  movel([-0.123614, -0.788371, -2.798725, -1.125292, 1.570796, 1.447182],accel_mss,speed_ms,0,blend_radius_m)
  movel([-0.122358, -0.787472, -2.798871, -1.126045, 1.570796, 1.448438],accel_mss,speed_ms,0,blend_radius_m)
  movel([-0.121105, -0.786979, -2.798951, -1.126459, 1.570796, 1.449692],accel_mss,speed_ms,0,blend_radius_m)
  movel([-0.120159, -0.787158, -2.798922, -1.126309, 1.570796, 1.450637],accel_mss,speed_ms,0,blend_radius_m)
  movel([-0.119008, -0.788690, -2.798674, -1.125025, 1.570796, 1.451789],accel_mss,speed_ms,0,blend_radius_m)
  movel([-0.118135, -0.791492, -2.798216, -1.122680, 1.570796, 1.452661],accel_mss,speed_ms,0,blend_radius_m)
  movel([-0.117601, -0.794594, -2.797706, -1.120090, 1.570796, 1.453195],accel_mss,speed_ms,0,blend_radius_m)
  movel([-0.115239, -0.789926, -2.798473, -1.123991, 1.570796, 1.455558],accel_mss,speed_ms,0,blend_radius_m)
  movel([-0.112520, -0.785198, -2.799238, -1.127953, 1.570796, 1.458276],accel_mss,speed_ms,0,blend_radius_m)
  movel([-0.109499, -0.780473, -2.799992, -1.131924, 1.570796, 1.461298],accel_mss,speed_ms,0,blend_radius_m)
  movel([-0.106241, -0.775820, -2.800723, -1.135846, 1.570796, 1.464556],accel_mss,speed_ms,0,blend_radius_m)
  movel([-0.099689, -0.766469, -2.802160, -1.143759, 1.570796, 1.471108],accel_mss,speed_ms,0,blend_radius_m)
  movel([-0.097728, -0.763893, -2.802549, -1.145948, 1.570796, 1.473068],accel_mss,speed_ms,0,blend_radius_m)
  movel([-0.095794, -0.761589, -2.802893, -1.147907, 1.570796, 1.475003],accel_mss,speed_ms,0,blend_radius_m)
  movel([-0.093954, -0.759736, -2.803169, -1.149484, 1.570796, 1.476842],accel_mss,speed_ms,0,blend_radius_m)
  movel([-0.092299, -0.758522, -2.803348, -1.150519, 1.570796, 1.478498],accel_mss,speed_ms,0,blend_radius_m)
  movel([-0.090884, -0.758158, -2.803402, -1.150829, 1.570796, 1.479912],accel_mss,speed_ms,0,blend_radius_m)
  movel([-0.089878, -0.758679, -2.803325, -1.150385, 1.570796, 1.480919],accel_mss,speed_ms,0,blend_radius_m)
  movel([-0.089251, -0.759892, -2.803145, -1.149351, 1.570796, 1.481545],accel_mss,speed_ms,0,blend_radius_m)
  movel([-0.088991, -0.761609, -2.802890, -1.147890, 1.570796, 1.481805],accel_mss,speed_ms,0,blend_radius_m)
  movel([-0.089073, -0.763633, -2.802588, -1.146168, 1.570796, 1.481724],accel_mss,speed_ms,0,blend_radius_m)
  movel([-0.089471, -0.765770, -2.802266, -1.144353, 1.570796, 1.481326],accel_mss,speed_ms,0,blend_radius_m)
  movel([-0.090165, -0.767829, -2.801954, -1.142606, 1.570796, 1.480631],accel_mss,speed_ms,0,blend_radius_m)
  movel([-0.091138, -0.769624, -2.801680, -1.141085, 1.570796, 1.479658],accel_mss,speed_ms,0,blend_radius_m)
  movel([-0.085055, -0.761341, -2.802930, -1.148118, 1.570796, 1.485742],accel_mss,speed_ms,0,blend_radius_m)
  movel([-0.081792, -0.757306, -2.803527, -1.151555, 1.570796, 1.489004],accel_mss,speed_ms,0,blend_radius_m)
  movel([-0.078396, -0.753391, -2.804099, -1.154899, 1.570796, 1.492400],accel_mss,speed_ms,0,blend_radius_m)
  movel([-0.074888, -0.749633, -2.804641, -1.158115, 1.570796, 1.495909],accel_mss,speed_ms,0,blend_radius_m)
  movel([-0.071275, -0.746070, -2.805148, -1.161171, 1.570796, 1.499521],accel_mss,speed_ms,0,blend_radius_m)
  movel([-0.067576, -0.742740, -2.805617, -1.164032, 1.570796, 1.503221],accel_mss,speed_ms,0,blend_radius_m)
  movel([-0.063806, -0.739679, -2.806043, -1.166667, 1.570796, 1.506991],accel_mss,speed_ms,0,blend_radius_m)
  movel([-0.061242, -0.738118, -2.806259, -1.168012, 1.570796, 1.509554],accel_mss,speed_ms,0,blend_radius_m)
  movel([-0.058496, -0.737145, -2.806393, -1.168852, 1.570796, 1.512301],accel_mss,speed_ms,0,blend_radius_m)
  movel([-0.057304, -0.737032, -2.806408, -1.168948, 1.570796, 1.513493],accel_mss,speed_ms,0,blend_radius_m)
  movel([-0.056360, -0.737246, -2.806379, -1.168764, 1.570796, 1.514437],accel_mss,speed_ms,0,blend_radius_m)
  movel([-0.055759, -0.737845, -2.806297, -1.168247, 1.570796, 1.515037],accel_mss,speed_ms,0,blend_radius_m)
  movel([-0.055607, -0.738896, -2.806152, -1.167342, 1.570796, 1.515190],accel_mss,speed_ms,0,blend_radius_m)
  movel([-0.055970, -0.740265, -2.805962, -1.166162, 1.570796, 1.514827],accel_mss,speed_ms,0,blend_radius_m)
  movel([-0.056714, -0.741799, -2.805748, -1.164841, 1.570796, 1.514083],accel_mss,speed_ms,0,blend_radius_m)
  movel([-0.058927, -0.745239, -2.805266, -1.161885, 1.570796, 1.511869],accel_mss,speed_ms,0,blend_radius_m)
  movel([-0.061573, -0.748454, -2.804809, -1.159126, 1.570796, 1.509223],accel_mss,speed_ms,0,blend_radius_m)
  movel([-0.064470, -0.751417, -2.804384, -1.156588, 1.570796, 1.506326],accel_mss,speed_ms,0,blend_radius_m)
  movel([-0.067437, -0.754102, -2.803995, -1.154291, 1.570796, 1.503359],accel_mss,speed_ms,0,blend_radius_m)
  movel([-0.063607, -0.752594, -2.804214, -1.155581, 1.570796, 1.507189],accel_mss,speed_ms,0,blend_radius_m)
  movel([-0.059620, -0.750631, -2.804497, -1.157260, 1.570796, 1.511176],accel_mss,speed_ms,0,blend_radius_m)
  movel([-0.055519, -0.748238, -2.804840, -1.159311, 1.570796, 1.515278],accel_mss,speed_ms,0,blend_radius_m)
  movel([-0.051338, -0.745435, -2.805238, -1.161716, 1.570796, 1.519459],accel_mss,speed_ms,0,blend_radius_m)
  movel([-0.048030, -0.742875, -2.805598, -1.163916, 1.570796, 1.522766],accel_mss,speed_ms,0,blend_radius_m)
  movel([-0.041537, -0.737330, -2.806367, -1.168691, 1.570796, 1.529259],accel_mss,speed_ms,0,blend_radius_m)
  movel([-0.038202, -0.734723, -2.806724, -1.170942, 1.570796, 1.532595],accel_mss,speed_ms,0,blend_radius_m)
  movel([-0.034400, -0.732028, -2.807090, -1.173271, 1.570796, 1.536396],accel_mss,speed_ms,0,blend_radius_m)
  movel([-0.027997, -0.727831, -2.807652, -1.176906, 1.570796, 1.542799],accel_mss,speed_ms,0,blend_radius_m)
  movel([-0.024935, -0.726094, -2.807883, -1.178413, 1.570796, 1.545861],accel_mss,speed_ms,0,blend_radius_m)
  movel([-0.022568, -0.725095, -2.808015, -1.179280, 1.570796, 1.548229],accel_mss,speed_ms,0,blend_radius_m)
  movel([-0.021784, -0.724985, -2.808029, -1.179375, 1.570796, 1.549013],accel_mss,speed_ms,0,blend_radius_m)
  movel([-0.021347, -0.725203, -2.808001, -1.179186, 1.570796, 1.549449],accel_mss,speed_ms,0,blend_radius_m)
  movel([-0.021306, -0.725781, -2.807924, -1.178683, 1.570796, 1.549490],accel_mss,speed_ms,0,blend_radius_m)
  movel([-0.021722, -0.726772, -2.807793, -1.177824, 1.570796, 1.549074],accel_mss,speed_ms,0,blend_radius_m)
  movel([-0.023301, -0.729254, -2.807462, -1.175672, 1.570796, 1.547495],accel_mss,speed_ms,0,blend_radius_m)
  movel([-0.025347, -0.731856, -2.807113, -1.173420, 1.570796, 1.545450],accel_mss,speed_ms,0,blend_radius_m)
  movel([-0.027725, -0.734514, -2.806753, -1.171123, 1.570796, 1.543072],accel_mss,speed_ms,0,blend_radius_m)
  movel([-0.030292, -0.737144, -2.806393, -1.168852, 1.570796, 1.540504],accel_mss,speed_ms,0,blend_radius_m)
  movel([-0.035478, -0.742049, -2.805713, -1.164626, 1.570796, 1.535318],accel_mss,speed_ms,0,blend_radius_m)
  movel([-0.039835, -0.745995, -2.805159, -1.161235, 1.570796, 1.530962],accel_mss,speed_ms,0,blend_radius_m)
  movel([-0.037640, -0.745598, -2.805215, -1.161576, 1.570796, 1.533156],accel_mss,speed_ms,0,blend_radius_m)
  movel([-0.035326, -0.744930, -2.805309, -1.162150, 1.570796, 1.535470],accel_mss,speed_ms,0,blend_radius_m)
  movel([-0.030418, -0.742923, -2.805591, -1.163875, 1.570796, 1.540378],accel_mss,speed_ms,0,blend_radius_m)
  movel([-0.025249, -0.740229, -2.805967, -1.166193, 1.570796, 1.545548],accel_mss,speed_ms,0,blend_radius_m)
  movel([-0.019955, -0.737110, -2.806398, -1.168881, 1.570796, 1.550841],accel_mss,speed_ms,0,blend_radius_m)
  movel([-0.015550, -0.734257, -2.806788, -1.171345, 1.570796, 1.555246],accel_mss,speed_ms,0,blend_radius_m)
  movel([-0.002182, -0.725105, -2.808013, -1.179270, 1.570796, 1.568614],accel_mss,speed_ms,0,blend_radius_m)
  movel([0.000291, -0.723828, -2.808181, -1.180380, 1.570796, 1.571087],accel_mss,speed_ms,0,blend_radius_m)
  movel([0.002219, -0.723407, -2.808237, -1.180746, 1.570796, 1.573015],accel_mss,speed_ms,0,blend_radius_m)
  movel([0.002614, -0.723722, -2.808195, -1.180471, 1.570796, 1.573410],accel_mss,speed_ms,0,blend_radius_m)
  movel([0.002432, -0.724499, -2.808093, -1.179796, 1.570796, 1.573228],accel_mss,speed_ms,0,blend_radius_m)
  movel([0.001528, -0.725818, -2.807919, -1.178652, 1.570796, 1.572325],accel_mss,speed_ms,0,blend_radius_m)
  movel([-0.000242, -0.727756, -2.807662, -1.176971, 1.570796, 1.570554],accel_mss,speed_ms,0,blend_radius_m)
  movel([-0.003204, -0.730567, -2.807287, -1.174536, 1.570796, 1.567592],accel_mss,speed_ms,0,blend_radius_m)
  movel([-0.006618, -0.733453, -2.806897, -1.172039, 1.570796, 1.564179],accel_mss,speed_ms,0,blend_radius_m)
  movel([-0.009977, -0.735885, -2.806566, -1.169939, 1.570796, 1.560819],accel_mss,speed_ms,0,blend_radius_m)
  movel([-0.011482, -0.736767, -2.806445, -1.169177, 1.570796, 1.559315],accel_mss,speed_ms,0,blend_radius_m)
  movel([-0.012779, -0.737329, -2.806368, -1.168692, 1.570796, 1.558017],accel_mss,speed_ms,0,blend_radius_m)
  movel([-0.007737, -0.737133, -2.806395, -1.168862, 1.570796, 1.563059],accel_mss,speed_ms,0,blend_radius_m)
  movel([-0.002332, -0.736239, -2.806517, -1.169632, 1.570796, 1.568464],accel_mss,speed_ms,0,blend_radius_m)
  movel([0.003362, -0.734781, -2.806716, -1.170892, 1.570796, 1.574158],accel_mss,speed_ms,0,blend_radius_m)
  movel([0.009278, -0.732894, -2.806973, -1.172522, 1.570796, 1.580074],accel_mss,speed_ms,0,blend_radius_m)
  movel([0.021466, -0.728361, -2.807582, -1.176446, 1.570796, 1.592262],accel_mss,speed_ms,0,blend_radius_m)
  movel([0.033600, -0.723736, -2.808193, -1.180459, 1.570796, 1.604396],accel_mss,speed_ms,0,blend_radius_m)
  movel([0.035605, -0.723312, -2.808249, -1.180828, 1.570796, 1.606402],accel_mss,speed_ms,0,blend_radius_m)
  movel([0.036255, -0.723590, -2.808212, -1.180586, 1.570796, 1.607051],accel_mss,speed_ms,0,blend_radius_m)
  movel([0.036422, -0.724403, -2.808106, -1.179880, 1.570796, 1.607218],accel_mss,speed_ms,0,blend_radius_m)
  movel([0.036036, -0.725600, -2.807948, -1.178841, 1.570796, 1.606833],accel_mss,speed_ms,0,blend_radius_m)
  movel([0.034004, -0.728911, -2.807508, -1.175970, 1.570796, 1.604800],accel_mss,speed_ms,0,blend_radius_m)
  movel([0.032557, -0.730811, -2.807254, -1.174324, 1.570796, 1.603354],accel_mss,speed_ms,0,blend_radius_m)
  movel([0.029315, -0.734343, -2.806776, -1.171270, 1.570796, 1.600111],accel_mss,speed_ms,0,blend_radius_m)
  movel([0.025758, -0.737485, -2.806346, -1.168557, 1.570796, 1.596555],accel_mss,speed_ms,0,blend_radius_m)
  movel([0.022037, -0.740240, -2.805965, -1.166184, 1.570796, 1.592834],accel_mss,speed_ms,0,blend_radius_m)
  movel([0.018315, -0.742582, -2.805639, -1.164168, 1.570796, 1.589112],accel_mss,speed_ms,0,blend_radius_m)
  movel([0.014745, -0.744506, -2.805369, -1.162514, 1.570796, 1.585541],accel_mss,speed_ms,0,blend_radius_m)
  movel([0.011481, -0.745991, -2.805159, -1.161239, 1.570796, 1.582277],accel_mss,speed_ms,0,blend_radius_m)
  movel([0.008687, -0.747012, -2.805015, -1.160363, 1.570796, 1.579483],accel_mss,speed_ms,0,blend_radius_m)
  movel([0.008653, -0.747858, -2.804894, -1.159637, 1.570796, 1.579449],accel_mss,speed_ms,0,blend_radius_m)
  movel([0.009139, -0.748262, -2.804836, -1.159290, 1.570796, 1.579935],accel_mss,speed_ms,0,blend_radius_m)
  movel([0.010647, -0.748657, -2.804780, -1.158952, 1.570796, 1.581444],accel_mss,speed_ms,0,blend_radius_m)
  movel([0.012360, -0.748723, -2.804771, -1.158895, 1.570796, 1.583157],accel_mss,speed_ms,0,blend_radius_m)
  movel([0.016128, -0.748272, -2.804835, -1.159282, 1.570796, 1.586925],accel_mss,speed_ms,0,blend_radius_m)
  movel([0.022850, -0.747039, -2.805011, -1.160339, 1.570796, 1.593647],accel_mss,speed_ms,0,blend_radius_m)
  movel([0.029687, -0.745518, -2.805226, -1.161645, 1.570796, 1.600483],accel_mss,speed_ms,0,blend_radius_m)
  movel([0.043712, -0.741725, -2.805759, -1.164905, 1.570796, 1.614508],accel_mss,speed_ms,0,blend_radius_m)
  movel([0.047601, -0.740757, -2.805894, -1.165738, 1.570796, 1.618397],accel_mss,speed_ms,0,blend_radius_m)
  movel([0.050057, -0.740378, -2.805946, -1.166065, 1.570796, 1.620854],accel_mss,speed_ms,0,blend_radius_m)
  movel([0.052405, -0.740305, -2.805956, -1.166128, 1.570796, 1.623201],accel_mss,speed_ms,0,blend_radius_m)
  movel([0.054288, -0.740724, -2.805898, -1.165767, 1.570796, 1.625084],accel_mss,speed_ms,0,blend_radius_m)
  movel([0.055366, -0.741799, -2.805748, -1.164841, 1.570796, 1.626162],accel_mss,speed_ms,0,blend_radius_m)
  movel([0.055503, -0.742631, -2.805632, -1.164126, 1.570796, 1.626300],accel_mss,speed_ms,0,blend_radius_m)
  movel([0.055317, -0.743690, -2.805484, -1.163216, 1.570796, 1.626113],accel_mss,speed_ms,0,blend_radius_m)
  movel([0.054755, -0.745002, -2.805299, -1.162088, 1.570796, 1.625552],accel_mss,speed_ms,0,blend_radius_m)
  movel([0.053791, -0.746577, -2.805076, -1.160736, 1.570796, 1.624588],accel_mss,speed_ms,0,blend_radius_m)
  movel([0.052380, -0.748019, -2.804871, -1.159499, 1.570796, 1.623176],accel_mss,speed_ms,0,blend_radius_m)
  movel([0.050460, -0.749382, -2.804676, -1.158330, 1.570796, 1.621256],accel_mss,speed_ms,0,blend_radius_m)
  movel([0.040183, -0.755535, -2.803787, -1.153068, 1.570796, 1.610979],accel_mss,speed_ms,0,blend_radius_m)
  movel([0.036738, -0.757148, -2.803550, -1.151690, 1.570796, 1.607535],accel_mss,speed_ms,0,blend_radius_m)
  movel([0.035260, -0.757597, -2.803484, -1.151307, 1.570796, 1.606056],accel_mss,speed_ms,0,blend_radius_m)
  movel([0.034042, -0.757700, -2.803469, -1.151220, 1.570796, 1.604838],accel_mss,speed_ms,0,blend_radius_m)
  movel([0.039097, -0.759244, -2.803241, -1.149904, 1.570796, 1.609893],accel_mss,speed_ms,0,blend_radius_m)
  movel([0.044720, -0.759886, -2.803146, -1.149356, 1.570796, 1.615516],accel_mss,speed_ms,0,blend_radius_m)
  movel([0.050778, -0.759793, -2.803160, -1.149436, 1.570796, 1.621574],accel_mss,speed_ms,0,blend_radius_m)
  movel([0.057144, -0.759117, -2.803260, -1.150012, 1.570796, 1.627940],accel_mss,speed_ms,0,blend_radius_m)
  movel([0.062648, -0.757727, -2.803465, -1.151197, 1.570796, 1.633444],accel_mss,speed_ms,0,blend_radius_m)
  movel([0.070534, -0.755900, -2.803733, -1.152756, 1.570796, 1.641330],accel_mss,speed_ms,0,blend_radius_m)
  movel([0.074102, -0.755520, -2.803789, -1.153080, 1.570796, 1.644899],accel_mss,speed_ms,0,blend_radius_m)
  movel([0.076754, -0.755848, -2.803741, -1.152800, 1.570796, 1.647550],accel_mss,speed_ms,0,blend_radius_m)
  movel([0.077577, -0.756361, -2.803666, -1.152363, 1.570796, 1.648374],accel_mss,speed_ms,0,blend_radius_m)
  movel([0.077981, -0.757146, -2.803551, -1.151692, 1.570796, 1.648777],accel_mss,speed_ms,0,blend_radius_m)
  movel([0.077904, -0.758242, -2.803389, -1.150758, 1.570796, 1.648701],accel_mss,speed_ms,0,blend_radius_m)
  movel([0.077296, -0.759666, -2.803179, -1.149544, 1.570796, 1.648093],accel_mss,speed_ms,0,blend_radius_m)
  movel([0.076368, -0.761124, -2.802963, -1.148302, 1.570796, 1.647164],accel_mss,speed_ms,0,blend_radius_m)
  movel([0.075295, -0.762513, -2.802755, -1.147120, 1.570796, 1.646091],accel_mss,speed_ms,0,blend_radius_m)
  movel([0.072924, -0.765097, -2.802368, -1.144925, 1.570796, 1.643720],accel_mss,speed_ms,0,blend_radius_m)
  movel([0.070302, -0.767643, -2.801982, -1.142764, 1.570796, 1.641099],accel_mss,speed_ms,0,blend_radius_m)
  movel([0.064988, -0.772160, -2.801291, -1.138938, 1.570796, 1.635784],accel_mss,speed_ms,0,blend_radius_m)
  movel([0.062326, -0.774111, -2.800989, -1.137289, 1.570796, 1.633122],accel_mss,speed_ms,0,blend_radius_m)
  movel([0.067181, -0.773517, -2.801081, -1.137791, 1.570796, 1.637977],accel_mss,speed_ms,0,blend_radius_m)
  movel([0.072189, -0.772546, -2.801231, -1.138612, 1.570796, 1.642985],accel_mss,speed_ms,0,blend_radius_m)
  movel([0.077338, -0.771243, -2.801432, -1.139714, 1.570796, 1.648134],accel_mss,speed_ms,0,blend_radius_m)
  movel([0.082615, -0.769641, -2.801678, -1.141070, 1.570796, 1.653412],accel_mss,speed_ms,0,blend_radius_m)
  movel([0.093490, -0.765710, -2.802275, -1.144404, 1.570796, 1.664286],accel_mss,speed_ms,0,blend_radius_m)
  movel([0.104701, -0.761055, -2.802973, -1.148361, 1.570796, 1.675497],accel_mss,speed_ms,0,blend_radius_m)
  movel([0.107639, -0.760148, -2.803108, -1.149134, 1.570796, 1.678435],accel_mss,speed_ms,0,blend_radius_m)
  movel([0.108683, -0.760339, -2.803079, -1.148971, 1.570796, 1.679480],accel_mss,speed_ms,0,blend_radius_m)
  movel([0.109107, -0.761285, -2.802939, -1.148165, 1.570796, 1.679903],accel_mss,speed_ms,0,blend_radius_m)
  movel([0.108974, -0.762254, -2.802794, -1.147340, 1.570796, 1.679770],accel_mss,speed_ms,0,blend_radius_m)
  movel([0.108569, -0.763342, -2.802631, -1.146416, 1.570796, 1.679365],accel_mss,speed_ms,0,blend_radius_m)
  movel([0.107060, -0.765815, -2.802259, -1.144315, 1.570796, 1.677856],accel_mss,speed_ms,0,blend_radius_m)
  movel([0.104857, -0.768511, -2.801850, -1.142028, 1.570796, 1.675653],accel_mss,speed_ms,0,blend_radius_m)
  movel([0.102226, -0.771265, -2.801429, -1.139696, 1.570796, 1.673022],accel_mss,speed_ms,0,blend_radius_m)
  movel([0.096762, -0.776227, -2.800659, -1.135502, 1.570796, 1.667558],accel_mss,speed_ms,0,blend_radius_m)
  movel([0.092780, -0.779303, -2.800177, -1.132910, 1.570796, 1.663577],accel_mss,speed_ms,0,blend_radius_m)
  movel([0.095018, -0.778629, -2.800283, -1.133477, 1.570796, 1.665815],accel_mss,speed_ms,0,blend_radius_m)
  movel([0.097342, -0.777697, -2.800429, -1.134262, 1.570796, 1.668138],accel_mss,speed_ms,0,blend_radius_m)
  movel([0.102193, -0.775141, -2.800829, -1.136419, 1.570796, 1.672990],accel_mss,speed_ms,0,blend_radius_m)
  movel([0.107238, -0.771741, -2.801355, -1.139293, 1.570796, 1.678035],accel_mss,speed_ms,0,blend_radius_m)
  movel([0.112383, -0.767625, -2.801985, -1.142779, 1.570796, 1.683179],accel_mss,speed_ms,0,blend_radius_m)
  movel([0.117534, -0.762890, -2.802699, -1.146800, 1.570796, 1.688330],accel_mss,speed_ms,0,blend_radius_m)
  movel([0.122590, -0.757669, -2.803474, -1.151246, 1.570796, 1.693387],accel_mss,speed_ms,0,blend_radius_m)
  movel([0.127452, -0.752066, -2.804291, -1.156033, 1.570796, 1.698249],accel_mss,speed_ms,0,blend_radius_m)
  movel([0.132018, -0.746209, -2.805128, -1.161051, 1.570796, 1.702814],accel_mss,speed_ms,0,blend_radius_m)
  movel([0.134037, -0.743591, -2.805498, -1.163300, 1.570796, 1.704834],accel_mss,speed_ms,0,blend_radius_m)
  movel([0.135120, -0.742450, -2.805657, -1.164281, 1.570796, 1.705916],accel_mss,speed_ms,0,blend_radius_m)
  movel([0.136237, -0.741570, -2.805780, -1.165038, 1.570796, 1.707033],accel_mss,speed_ms,0,blend_radius_m)
  movel([0.137379, -0.741088, -2.805848, -1.165453, 1.570796, 1.708175],accel_mss,speed_ms,0,blend_radius_m)
  movel([0.138333, -0.741050, -2.805853, -1.165486, 1.570796, 1.709129],accel_mss,speed_ms,0,blend_radius_m)
  movel([0.139345, -0.741714, -2.805760, -1.164914, 1.570796, 1.710141],accel_mss,speed_ms,0,blend_radius_m)
  movel([0.139829, -0.743141, -2.805561, -1.163688, 1.570796, 1.710625],accel_mss,speed_ms,0,blend_radius_m)
  movel([0.139879, -0.745135, -2.805280, -1.161974, 1.570796, 1.710675],accel_mss,speed_ms,0,blend_radius_m)
  movel([0.139591, -0.747520, -2.804942, -1.159927, 1.570796, 1.710387],accel_mss,speed_ms,0,blend_radius_m)
  movel([0.138373, -0.752698, -2.804199, -1.155492, 1.570796, 1.709169],accel_mss,speed_ms,0,blend_radius_m)
  movel([0.136926, -0.757207, -2.803542, -1.151641, 1.570796, 1.707723],accel_mss,speed_ms,0,blend_radius_m)
  movel([0.140852, -0.751503, -2.804372, -1.156514, 1.570796, 1.711648],accel_mss,speed_ms,0,blend_radius_m)
  movel([0.144402, -0.745687, -2.805202, -1.161500, 1.570796, 1.715198],accel_mss,speed_ms,0,blend_radius_m)
  movel([0.147549, -0.739819, -2.806024, -1.166546, 1.570796, 1.718345],accel_mss,speed_ms,0,blend_radius_m)
  movel([0.150273, -0.733978, -2.806826, -1.171585, 1.570796, 1.721070],accel_mss,speed_ms,0,blend_radius_m)
  movel([0.152533, -0.728242, -2.807598, -1.176549, 1.570796, 1.723330],accel_mss,speed_ms,0,blend_radius_m)
  movel([0.154318, -0.722674, -2.808332, -1.181382, 1.570796, 1.725114],accel_mss,speed_ms,0,blend_radius_m)
  movel([0.155580, -0.717372, -2.809019, -1.185998, 1.570796, 1.726376],accel_mss,speed_ms,0,blend_radius_m)
  movel([0.156297, -0.712407, -2.809651, -1.190332, 1.570796, 1.727094],accel_mss,speed_ms,0,blend_radius_m)
  movel([0.156402, -0.706121, -2.810434, -1.195834, 1.570796, 1.727198],accel_mss,speed_ms,0,blend_radius_m)
  movel([0.156716, -0.702641, -2.810860, -1.198888, 1.570796, 1.727512],accel_mss,speed_ms,0,blend_radius_m)
  movel([0.157110, -0.700860, -2.811076, -1.200453, 1.570796, 1.727906],accel_mss,speed_ms,0,blend_radius_m)
  movel([0.157721, -0.699072, -2.811292, -1.202026, 1.570796, 1.728517],accel_mss,speed_ms,0,blend_radius_m)
  movel([0.159157, -0.696129, -2.811643, -1.204617, 1.570796, 1.729953],accel_mss,speed_ms,0,blend_radius_m)
  movel([0.160486, -0.694322, -2.811857, -1.206209, 1.570796, 1.731283],accel_mss,speed_ms,0,blend_radius_m)
  movel([0.161725, -0.693413, -2.811965, -1.207012, 1.570796, 1.732521],accel_mss,speed_ms,0,blend_radius_m)
  movel([0.162880, -0.693157, -2.811995, -1.207237, 1.570796, 1.733676],accel_mss,speed_ms,0,blend_radius_m)
  movel([0.165920, -0.693920, -2.811905, -1.206564, 1.570796, 1.736716],accel_mss,speed_ms,0,blend_radius_m)
  movel([0.166833, -0.693867, -2.811911, -1.206611, 1.570796, 1.737629],accel_mss,speed_ms,0,blend_radius_m)
  movel([0.168876, -0.689499, -2.812422, -1.210468, 1.570796, 1.739672],accel_mss,speed_ms,0,blend_radius_m)
  movel([0.170617, -0.685171, -2.812919, -1.214299, 1.570796, 1.741413],accel_mss,speed_ms,0,blend_radius_m)
  movel([0.172069, -0.680901, -2.813402, -1.218086, 1.570796, 1.742866],accel_mss,speed_ms,0,blend_radius_m)
  movel([0.173248, -0.676699, -2.813870, -1.221820, 1.570796, 1.744044],accel_mss,speed_ms,0,blend_radius_m)
  movel([0.174153, -0.672593, -2.814320, -1.225476, 1.570796, 1.744950],accel_mss,speed_ms,0,blend_radius_m)
  movel([0.174801, -0.668595, -2.814751, -1.229043, 1.570796, 1.745598],accel_mss,speed_ms,0,blend_radius_m)
  movel([0.175391, -0.660973, -2.815554, -1.235862, 1.570796, 1.746188],accel_mss,speed_ms,0,blend_radius_m)
  movel([0.175103, -0.653985, -2.816269, -1.242134, 1.570796, 1.745899],accel_mss,speed_ms,0,blend_radius_m)
  movel([0.174059, -0.647747, -2.816891, -1.247751, 1.570796, 1.744855],accel_mss,speed_ms,0,blend_radius_m)
  movel([0.172351, -0.642405, -2.817410, -1.252574, 1.570796, 1.743147],accel_mss,speed_ms,0,blend_radius_m)
  movel([0.170116, -0.638064, -2.817824, -1.256502, 1.570796, 1.740912],accel_mss,speed_ms,0,blend_radius_m)
  speed_ms = 0.005
  movel([0.170116, -0.631907, -2.811057, -1.269425, 1.570796, 1.740912],accel_mss,speed_ms,0,blend_radius_m)
  speed_ms = 0.040
  movel([0.138700, -0.656581, -2.808612, -1.247195, 1.570796, 1.709497],accel_mss,speed_ms,0,blend_radius_m)
  speed_ms = 0.005
  movel([0.138700, -0.663123, -2.815330, -1.233936, 1.570796, 1.709497],accel_mss,speed_ms,0,blend_radius_m)
  speed_ms = 0.025
  movel([0.136102, -0.662756, -2.815369, -1.234264, 1.570796, 1.706899],accel_mss,speed_ms,0,blend_radius_m)
  movel([0.133054, -0.663285, -2.815313, -1.233791, 1.570796, 1.703850],accel_mss,speed_ms,0,blend_radius_m)
  movel([0.129644, -0.664578, -2.815178, -1.232634, 1.570796, 1.700441],accel_mss,speed_ms,0,blend_radius_m)
  movel([0.125976, -0.666489, -2.814975, -1.230924, 1.570796, 1.696772],accel_mss,speed_ms,0,blend_radius_m)
  movel([0.122143, -0.668882, -2.814720, -1.228787, 1.570796, 1.692939],accel_mss,speed_ms,0,blend_radius_m)
  movel([0.118234, -0.671617, -2.814426, -1.226346, 1.570796, 1.689030],accel_mss,speed_ms,0,blend_radius_m)
  movel([0.110564, -0.677562, -2.813775, -1.221052, 1.570796, 1.681360],accel_mss,speed_ms,0,blend_radius_m)
  speed_ms = 0.005
  movel([0.110564, -0.670808, -2.807087, -1.234494, 1.570796, 1.681360],accel_mss,speed_ms,0,blend_radius_m)
  speed_ms = 0.040
  movel([0.120496, -0.662365, -2.808003, -1.242021, 1.570796, 1.691293],accel_mss,speed_ms,0,blend_radius_m)
  speed_ms = 0.005
  movel([0.120496, -0.668994, -2.814708, -1.228687, 1.570796, 1.691293],accel_mss,speed_ms,0,blend_radius_m)
  speed_ms = 0.025
  movel([0.122110, -0.664213, -2.815216, -1.232960, 1.570796, 1.692907],accel_mss,speed_ms,0,blend_radius_m)
  movel([0.123299, -0.659769, -2.815679, -1.236941, 1.570796, 1.694095],accel_mss,speed_ms,0,blend_radius_m)
  movel([0.124068, -0.655656, -2.816100, -1.240632, 1.570796, 1.694864],accel_mss,speed_ms,0,blend_radius_m)
  movel([0.124435, -0.651859, -2.816483, -1.244047, 1.570796, 1.695231],accel_mss,speed_ms,0,blend_radius_m)
  movel([0.124423, -0.648357, -2.816831, -1.247202, 1.570796, 1.695219],accel_mss,speed_ms,0,blend_radius_m)
  movel([0.124046, -0.645138, -2.817146, -1.250105, 1.570796, 1.694842],accel_mss,speed_ms,0,blend_radius_m)
  movel([0.123323, -0.642185, -2.817431, -1.252773, 1.570796, 1.694119],accel_mss,speed_ms,0,blend_radius_m)
  movel([0.122274, -0.639481, -2.817690, -1.255219, 1.570796, 1.693071],accel_mss,speed_ms,0,blend_radius_m)
  movel([0.118229, -0.632565, -2.818336, -1.261487, 1.570796, 1.689025],accel_mss,speed_ms,0,blend_radius_m)
  movel([0.116481, -0.629055, -2.818657, -1.264676, 1.570796, 1.687277],accel_mss,speed_ms,0,blend_radius_m)
  movel([0.115290, -0.624496, -2.819067, -1.268826, 1.570796, 1.686086],accel_mss,speed_ms,0,blend_radius_m)
  movel([0.114590, -0.618038, -2.819633, -1.274718, 1.570796, 1.685386],accel_mss,speed_ms,0,blend_radius_m)
  movel([0.114549, -0.610974, -2.820233, -1.281182, 1.570796, 1.685345],accel_mss,speed_ms,0,blend_radius_m)
  movel([0.115398, -0.603180, -2.820873, -1.288336, 1.570796, 1.686195],accel_mss,speed_ms,0,blend_radius_m)
  movel([0.116229, -0.598970, -2.821209, -1.292210, 1.570796, 1.687025],accel_mss,speed_ms,0,blend_radius_m)
  movel([0.117376, -0.594532, -2.821555, -1.296302, 1.570796, 1.688172],accel_mss,speed_ms,0,blend_radius_m)
  movel([0.119840, -0.587296, -2.822104, -1.302989, 1.570796, 1.690636],accel_mss,speed_ms,0,blend_radius_m)
  movel([0.123098, -0.579856, -2.822647, -1.309886, 1.570796, 1.693894],accel_mss,speed_ms,0,blend_radius_m)
  movel([0.127112, -0.572263, -2.823180, -1.316946, 1.570796, 1.697908],accel_mss,speed_ms,0,blend_radius_m)
  movel([0.131842, -0.564581, -2.823697, -1.324111, 1.570796, 1.702638],accel_mss,speed_ms,0,blend_radius_m)
  movel([0.137234, -0.556886, -2.824193, -1.331309, 1.570796, 1.708030],accel_mss,speed_ms,0,blend_radius_m)
  movel([0.143247, -0.549247, -2.824664, -1.338478, 1.570796, 1.714044],accel_mss,speed_ms,0,blend_radius_m)
  movel([0.149829, -0.541732, -2.825106, -1.345550, 1.570796, 1.720625],accel_mss,speed_ms,0,blend_radius_m)
  movel([0.156913, -0.534435, -2.825516, -1.352438, 1.570796, 1.727709],accel_mss,speed_ms,0,blend_radius_m)
  movel([0.162439, -0.529240, -2.825796, -1.357352, 1.570796, 1.733235],accel_mss,speed_ms,0,blend_radius_m)
  movel([0.168059, -0.524374, -2.826050, -1.361965, 1.570796, 1.738855],accel_mss,speed_ms,0,blend_radius_m)
  movel([0.173713, -0.519879, -2.826276, -1.366234, 1.570796, 1.744510],accel_mss,speed_ms,0,blend_radius_m)
  movel([0.179359, -0.515772, -2.826477, -1.370140, 1.570796, 1.750155],accel_mss,speed_ms,0,blend_radius_m)
  movel([0.184932, -0.512108, -2.826651, -1.373629, 1.570796, 1.755728],accel_mss,speed_ms,0,blend_radius_m)
  movel([0.190379, -0.508915, -2.826799, -1.376675, 1.570796, 1.761175],accel_mss,speed_ms,0,blend_radius_m)
  movel([0.195640, -0.506227, -2.826921, -1.379241, 1.570796, 1.766437],accel_mss,speed_ms,0,blend_radius_m)
  movel([0.200660, -0.504082, -2.827016, -1.381291, 1.570796, 1.771456],accel_mss,speed_ms,0,blend_radius_m)
  movel([0.205378, -0.502513, -2.827085, -1.382791, 1.570796, 1.776175],accel_mss,speed_ms,0,blend_radius_m)
  movel([0.209750, -0.501543, -2.827127, -1.383719, 1.570796, 1.780546],accel_mss,speed_ms,0,blend_radius_m)
  movel([0.213716, -0.501208, -2.827141, -1.384040, 1.570796, 1.784512],accel_mss,speed_ms,0,blend_radius_m)
  movel([0.217226, -0.501531, -2.827127, -1.383731, 1.570796, 1.788023],accel_mss,speed_ms,0,blend_radius_m)
  movel([0.220235, -0.502533, -2.827084, -1.382772, 1.570796, 1.791031],accel_mss,speed_ms,0,blend_radius_m)
  movel([0.222682, -0.504249, -2.827009, -1.381132, 1.570796, 1.793478],accel_mss,speed_ms,0,blend_radius_m)
  movel([0.224532, -0.506682, -2.826900, -1.378807, 1.570796, 1.795329],accel_mss,speed_ms,0,blend_radius_m)
  movel([0.225745, -0.509859, -2.826756, -1.375774, 1.570796, 1.796541],accel_mss,speed_ms,0,blend_radius_m)
  movel([0.226531, -0.514797, -2.826524, -1.371068, 1.570796, 1.797328],accel_mss,speed_ms,0,blend_radius_m)
  movel([0.226728, -0.520288, -2.826256, -1.365845, 1.570796, 1.797524],accel_mss,speed_ms,0,blend_radius_m)
  movel([0.226455, -0.526200, -2.825956, -1.360233, 1.570796, 1.797251],accel_mss,speed_ms,0,blend_radius_m)
  movel([0.225856, -0.532375, -2.825628, -1.354386, 1.570796, 1.796653],accel_mss,speed_ms,0,blend_radius_m)
  movel([0.223911, -0.546253, -2.824843, -1.341294, 1.570796, 1.794707],accel_mss,speed_ms,0,blend_radius_m)
  movel([0.221348, -0.560558, -2.823959, -1.327872, 1.570796, 1.792145],accel_mss,speed_ms,0,blend_radius_m)
  movel([0.218336, -0.575144, -2.822980, -1.314265, 1.570796, 1.789132],accel_mss,speed_ms,0,blend_radius_m)
  movel([0.215033, -0.589850, -2.821912, -1.300626, 1.570796, 1.785830],accel_mss,speed_ms,0,blend_radius_m)
  movel([0.201838, -0.647356, -2.816929, -1.248104, 1.570796, 1.772635],accel_mss,speed_ms,0,blend_radius_m)
  movel([0.196552, -0.674366, -2.814127, -1.223896, 1.570796, 1.767348],accel_mss,speed_ms,0,blend_radius_m)
  movel([0.194383, -0.687392, -2.812665, -1.212332, 1.570796, 1.765179],accel_mss,speed_ms,0,blend_radius_m)
  movel([0.192649, -0.699989, -2.811181, -1.201218, 1.570796, 1.763445],accel_mss,speed_ms,0,blend_radius_m)
  movel([0.191422, -0.712103, -2.809689, -1.190597, 1.570796, 1.762219],accel_mss,speed_ms,0,blend_radius_m)
  movel([0.190783, -0.723666, -2.808203, -1.180520, 1.570796, 1.761579],accel_mss,speed_ms,0,blend_radius_m)
  movel([0.190794, -0.734632, -2.806737, -1.171020, 1.570796, 1.761590],accel_mss,speed_ms,0,blend_radius_m)
  movel([0.191537, -0.744943, -2.805307, -1.162139, 1.570796, 1.762333],accel_mss,speed_ms,0,blend_radius_m)
  movel([0.192118, -0.748698, -2.804774, -1.158917, 1.570796, 1.762914],accel_mss,speed_ms,0,blend_radius_m)
  movel([0.193186, -0.751978, -2.804303, -1.156107, 1.570796, 1.763982],accel_mss,speed_ms,0,blend_radius_m)
  movel([0.194999, -0.754344, -2.803960, -1.154085, 1.570796, 1.765795],accel_mss,speed_ms,0,blend_radius_m)
  movel([0.196267, -0.755045, -2.803858, -1.153486, 1.570796, 1.767064],accel_mss,speed_ms,0,blend_radius_m)
  movel([0.197826, -0.755346, -2.803814, -1.153229, 1.570796, 1.768623],accel_mss,speed_ms,0,blend_radius_m)
  speed_ms = 0.005
  movel([0.197826, -0.747557, -2.797313, -1.167520, 1.570796, 1.768623],accel_mss,speed_ms,0,blend_radius_m)
  speed_ms = 0.040
  movel([0.166317, -0.709653, -2.802474, -1.200262, 1.570796, 1.737113],accel_mss,speed_ms,0,blend_radius_m)
  speed_ms = 0.005
  movel([0.166317, -0.716956, -2.809072, -1.186361, 1.570796, 1.737113],accel_mss,speed_ms,0,blend_radius_m)
  speed_ms = 0.025
  movel([0.165098, -0.718894, -2.808823, -1.184672, 1.570796, 1.735894],accel_mss,speed_ms,0,blend_radius_m)
  movel([0.164169, -0.720873, -2.808567, -1.182949, 1.570796, 1.734965],accel_mss,speed_ms,0,blend_radius_m)
  movel([0.163511, -0.722861, -2.808308, -1.181220, 1.570796, 1.734307],accel_mss,speed_ms,0,blend_radius_m)
  movel([0.163074, -0.724875, -2.808044, -1.179471, 1.570796, 1.733870],accel_mss,speed_ms,0,blend_radius_m)
  movel([0.162764, -0.728898, -2.807510, -1.175981, 1.570796, 1.733560],accel_mss,speed_ms,0,blend_radius_m)
  movel([0.162975, -0.732871, -2.806976, -1.172543, 1.570796, 1.733771],accel_mss,speed_ms,0,blend_radius_m)
  movel([0.164204, -0.743735, -2.805477, -1.163177, 1.570796, 1.735001],accel_mss,speed_ms,0,blend_radius_m)
  movel([0.163980, -0.746745, -2.805052, -1.160591, 1.570796, 1.734776],accel_mss,speed_ms,0,blend_radius_m)
  movel([0.163462, -0.748245, -2.804839, -1.159305, 1.570796, 1.734258],accel_mss,speed_ms,0,blend_radius_m)
  movel([0.162572, -0.749528, -2.804656, -1.158205, 1.570796, 1.733369],accel_mss,speed_ms,0,blend_radius_m)
  movel([0.161731, -0.750298, -2.804545, -1.157545, 1.570796, 1.732527],accel_mss,speed_ms,0,blend_radius_m)
  movel([0.160936, -0.750613, -2.804500, -1.157276, 1.570796, 1.731733],accel_mss,speed_ms,0,blend_radius_m)
  movel([0.160186, -0.750538, -2.804511, -1.157340, 1.570796, 1.730982],accel_mss,speed_ms,0,blend_radius_m)
  movel([0.158834, -0.749419, -2.804671, -1.158299, 1.570796, 1.729630],accel_mss,speed_ms,0,blend_radius_m)
  movel([0.157687, -0.747402, -2.804959, -1.160028, 1.570796, 1.728483],accel_mss,speed_ms,0,blend_radius_m)
  movel([0.156071, -0.742470, -2.805655, -1.164264, 1.570796, 1.726867],accel_mss,speed_ms,0,blend_radius_m)
  movel([0.155517, -0.739344, -2.806090, -1.166956, 1.570796, 1.726314],accel_mss,speed_ms,0,blend_radius_m)
  movel([0.153840, -0.744960, -2.805305, -1.162125, 1.570796, 1.724636],accel_mss,speed_ms,0,blend_radius_m)
  movel([0.152864, -0.750190, -2.804561, -1.157639, 1.570796, 1.723661],accel_mss,speed_ms,0,blend_radius_m)
  movel([0.152485, -0.755065, -2.803855, -1.153468, 1.570796, 1.723281],accel_mss,speed_ms,0,blend_radius_m)
  movel([0.152612, -0.759591, -2.803190, -1.149608, 1.570796, 1.723409],accel_mss,speed_ms,0,blend_radius_m)
  movel([0.153139, -0.763802, -2.802562, -1.146024, 1.570796, 1.723935],accel_mss,speed_ms,0,blend_radius_m)
  movel([0.153986, -0.767697, -2.801974, -1.142718, 1.570796, 1.724782],accel_mss,speed_ms,0,blend_radius_m)
  movel([0.156246, -0.774616, -2.800910, -1.136862, 1.570796, 1.727042],accel_mss,speed_ms,0,blend_radius_m)
  movel([0.156304, -0.776266, -2.800653, -1.135470, 1.570796, 1.727100],accel_mss,speed_ms,0,blend_radius_m)
  movel([0.155931, -0.777204, -2.800507, -1.134678, 1.570796, 1.726728],accel_mss,speed_ms,0,blend_radius_m)
  movel([0.155223, -0.778000, -2.800382, -1.134007, 1.570796, 1.726019],accel_mss,speed_ms,0,blend_radius_m)
  movel([0.154317, -0.778384, -2.800321, -1.133684, 1.570796, 1.725113],accel_mss,speed_ms,0,blend_radius_m)
  movel([0.152367, -0.778552, -2.800295, -1.133542, 1.570796, 1.723163],accel_mss,speed_ms,0,blend_radius_m)
  movel([0.150735, -0.778213, -2.800348, -1.133827, 1.570796, 1.721532],accel_mss,speed_ms,0,blend_radius_m)
  movel([0.149384, -0.777445, -2.800469, -1.134475, 1.570796, 1.720180],accel_mss,speed_ms,0,blend_radius_m)
  movel([0.148290, -0.776299, -2.800648, -1.135442, 1.570796, 1.719086],accel_mss,speed_ms,0,blend_radius_m)
  movel([0.146758, -0.773161, -2.801136, -1.138092, 1.570796, 1.717554],accel_mss,speed_ms,0,blend_radius_m)
  movel([0.145914, -0.769328, -2.801725, -1.141336, 1.570796, 1.716710],accel_mss,speed_ms,0,blend_radius_m)
  movel([0.145148, -0.778136, -2.800360, -1.133893, 1.570796, 1.715944],accel_mss,speed_ms,0,blend_radius_m)
  movel([0.145196, -0.782168, -2.799723, -1.130499, 1.570796, 1.715993],accel_mss,speed_ms,0,blend_radius_m)
  movel([0.145776, -0.785782, -2.799144, -1.127463, 1.570796, 1.716573],accel_mss,speed_ms,0,blend_radius_m)
  movel([0.146955, -0.788308, -2.798736, -1.125345, 1.570796, 1.717752],accel_mss,speed_ms,0,blend_radius_m)
  movel([0.150125, -0.792178, -2.798104, -1.122107, 1.570796, 1.720921],accel_mss,speed_ms,0,blend_radius_m)
  movel([0.151210, -0.794682, -2.797691, -1.120016, 1.570796, 1.722006],accel_mss,speed_ms,0,blend_radius_m)
  movel([0.151294, -0.795308, -2.797587, -1.119493, 1.570796, 1.722090],accel_mss,speed_ms,0,blend_radius_m)
  movel([0.151105, -0.796095, -2.797457, -1.118837, 1.570796, 1.721902],accel_mss,speed_ms,0,blend_radius_m)
  movel([0.150490, -0.796935, -2.797317, -1.118137, 1.570796, 1.721287],accel_mss,speed_ms,0,blend_radius_m)
  movel([0.149467, -0.797739, -2.797183, -1.117467, 1.570796, 1.720263],accel_mss,speed_ms,0,blend_radius_m)
  movel([0.146733, -0.799179, -2.796941, -1.116269, 1.570796, 1.717529],accel_mss,speed_ms,0,blend_radius_m)
  movel([0.142223, -0.800846, -2.796661, -1.114882, 1.570796, 1.713020],accel_mss,speed_ms,0,blend_radius_m)
  movel([0.142758, -0.803053, -2.796287, -1.113049, 1.570796, 1.713554],accel_mss,speed_ms,0,blend_radius_m)
  movel([0.143619, -0.805415, -2.795885, -1.111089, 1.570796, 1.714415],accel_mss,speed_ms,0,blend_radius_m)
  movel([0.144902, -0.807761, -2.795482, -1.109146, 1.570796, 1.715698],accel_mss,speed_ms,0,blend_radius_m)
  movel([0.146705, -0.809923, -2.795108, -1.107358, 1.570796, 1.717501],accel_mss,speed_ms,0,blend_radius_m)
  movel([0.152042, -0.812028, -2.794742, -1.105619, 1.570796, 1.722838],accel_mss,speed_ms,0,blend_radius_m)
  movel([0.154980, -0.813362, -2.794508, -1.104519, 1.570796, 1.725776],accel_mss,speed_ms,0,blend_radius_m)
  movel([0.155811, -0.814073, -2.794384, -1.103932, 1.570796, 1.726607],accel_mss,speed_ms,0,blend_radius_m)
  movel([0.155954, -0.814801, -2.794255, -1.103332, 1.570796, 1.726751],accel_mss,speed_ms,0,blend_radius_m)
  movel([0.155514, -0.815661, -2.794104, -1.102624, 1.570796, 1.726310],accel_mss,speed_ms,0,blend_radius_m)
  movel([0.154880, -0.816481, -2.793959, -1.101949, 1.570796, 1.725676],accel_mss,speed_ms,0,blend_radius_m)
  movel([0.153372, -0.817748, -2.793735, -1.100907, 1.570796, 1.724168],accel_mss,speed_ms,0,blend_radius_m)
  movel([0.152148, -0.818307, -2.793635, -1.100447, 1.570796, 1.722944],accel_mss,speed_ms,0,blend_radius_m)
  movel([0.150940, -0.818620, -2.793579, -1.100190, 1.570796, 1.721736],accel_mss,speed_ms,0,blend_radius_m)
  movel([0.148664, -0.819018, -2.793508, -1.099862, 1.570796, 1.719461],accel_mss,speed_ms,0,blend_radius_m)
  movel([0.149487, -0.821978, -2.792978, -1.097433, 1.570796, 1.720283],accel_mss,speed_ms,0,blend_radius_m)
  movel([0.150580, -0.824668, -2.792492, -1.095228, 1.570796, 1.721377],accel_mss,speed_ms,0,blend_radius_m)
  movel([0.151941, -0.827078, -2.792054, -1.093257, 1.570796, 1.722738],accel_mss,speed_ms,0,blend_radius_m)
  movel([0.153547, -0.829212, -2.791663, -1.091514, 1.570796, 1.724344],accel_mss,speed_ms,0,blend_radius_m)
  movel([0.155518, -0.830855, -2.791360, -1.090174, 1.570796, 1.726315],accel_mss,speed_ms,0,blend_radius_m)
  movel([0.157892, -0.831960, -2.791156, -1.089273, 1.570796, 1.728688],accel_mss,speed_ms,0,blend_radius_m)
  movel([0.163164, -0.833388, -2.790891, -1.088110, 1.570796, 1.733961],accel_mss,speed_ms,0,blend_radius_m)
  movel([0.164477, -0.834123, -2.790754, -1.087512, 1.570796, 1.735273],accel_mss,speed_ms,0,blend_radius_m)
  movel([0.164731, -0.834865, -2.790615, -1.086908, 1.570796, 1.735527],accel_mss,speed_ms,0,blend_radius_m)
  movel([0.164486, -0.835941, -2.790414, -1.086034, 1.570796, 1.735282],accel_mss,speed_ms,0,blend_radius_m)
  movel([0.163859, -0.836981, -2.790219, -1.085189, 1.570796, 1.734656],accel_mss,speed_ms,0,blend_radius_m)
  movel([0.163012, -0.837903, -2.790045, -1.084441, 1.570796, 1.733808],accel_mss,speed_ms,0,blend_radius_m)
  movel([0.161071, -0.839356, -2.789770, -1.083263, 1.570796, 1.731867],accel_mss,speed_ms,0,blend_radius_m)
  movel([0.158538, -0.840756, -2.789505, -1.082128, 1.570796, 1.729334],accel_mss,speed_ms,0,blend_radius_m)
  movel([0.156117, -0.841803, -2.789305, -1.081281, 1.570796, 1.726913],accel_mss,speed_ms,0,blend_radius_m)
  movel([0.153793, -0.842552, -2.789162, -1.080675, 1.570796, 1.724589],accel_mss,speed_ms,0,blend_radius_m)
  movel([0.151559, -0.843038, -2.789069, -1.080282, 1.570796, 1.722355],accel_mss,speed_ms,0,blend_radius_m)
  movel([0.152827, -0.845070, -2.788679, -1.078639, 1.570796, 1.723624],accel_mss,speed_ms,0,blend_radius_m)
  movel([0.154404, -0.846724, -2.788360, -1.077305, 1.570796, 1.725200],accel_mss,speed_ms,0,blend_radius_m)
  movel([0.156283, -0.847956, -2.788121, -1.076312, 1.570796, 1.727080],accel_mss,speed_ms,0,blend_radius_m)
  movel([0.158458, -0.848729, -2.787971, -1.075689, 1.570796, 1.729255],accel_mss,speed_ms,0,blend_radius_m)
  movel([0.160934, -0.848998, -2.787919, -1.075472, 1.570796, 1.731730],accel_mss,speed_ms,0,blend_radius_m)
  movel([0.163710, -0.848723, -2.787972, -1.075694, 1.570796, 1.734507],accel_mss,speed_ms,0,blend_radius_m)
  movel([0.166787, -0.847855, -2.788141, -1.076393, 1.570796, 1.737583],accel_mss,speed_ms,0,blend_radius_m)
  movel([0.170171, -0.846352, -2.788432, -1.077605, 1.570796, 1.740967],accel_mss,speed_ms,0,blend_radius_m)
  speed_ms = 0.005
  movel([0.170171, -0.837613, -2.782198, -1.092579, 1.570796, 1.740967],accel_mss,speed_ms,0,blend_radius_m)
  speed_ms = 0.040
  movel([0.185325, -0.814540, -2.786475, -1.111374, 1.570796, 1.756121],accel_mss,speed_ms,0,blend_radius_m)
  speed_ms = 0.005
  movel([0.185325, -0.823064, -2.792783, -1.096542, 1.570796, 1.756121],accel_mss,speed_ms,0,blend_radius_m)
  speed_ms = 0.025
  movel([0.179130, -0.822911, -2.792810, -1.096668, 1.570796, 1.749926],accel_mss,speed_ms,0,blend_radius_m)
  movel([0.176504, -0.822539, -2.792877, -1.096973, 1.570796, 1.747300],accel_mss,speed_ms,0,blend_radius_m)
  movel([0.174175, -0.821867, -2.792998, -1.097524, 1.570796, 1.744971],accel_mss,speed_ms,0,blend_radius_m)
  movel([0.172123, -0.820815, -2.793187, -1.098387, 1.570796, 1.742919],accel_mss,speed_ms,0,blend_radius_m)
  movel([0.170335, -0.819304, -2.793457, -1.099628, 1.570796, 1.741131],accel_mss,speed_ms,0,blend_radius_m)
  movel([0.168788, -0.817262, -2.793821, -1.101306, 1.570796, 1.739584],accel_mss,speed_ms,0,blend_radius_m)
  movel([0.167475, -0.814605, -2.794290, -1.103494, 1.570796, 1.738271],accel_mss,speed_ms,0,blend_radius_m)
  movel([0.165467, -0.808324, -2.795385, -1.108681, 1.570796, 1.736263],accel_mss,speed_ms,0,blend_radius_m)
  movel([0.164156, -0.801360, -2.796574, -1.114455, 1.570796, 1.734952],accel_mss,speed_ms,0,blend_radius_m)
  movel([0.163481, -0.793797, -2.797837, -1.120755, 1.570796, 1.734277],accel_mss,speed_ms,0,blend_radius_m)
  movel([0.163370, -0.785739, -2.799151, -1.127499, 1.570796, 1.734166],accel_mss,speed_ms,0,blend_radius_m)
  movel([0.163693, -0.778798, -2.800256, -1.133335, 1.570796, 1.734489],accel_mss,speed_ms,0,blend_radius_m)
  movel([0.164351, -0.771584, -2.801380, -1.139426, 1.570796, 1.735147],accel_mss,speed_ms,0,blend_radius_m)
  movel([0.166427, -0.756480, -2.803648, -1.152261, 1.570796, 1.737223],accel_mss,speed_ms,0,blend_radius_m)
  movel([0.175526, -0.702006, -2.810937, -1.199445, 1.570796, 1.746322],accel_mss,speed_ms,0,blend_radius_m)
  movel([0.177448, -0.690287, -2.812330, -1.209772, 1.570796, 1.748244],accel_mss,speed_ms,0,blend_radius_m)
  movel([0.179180, -0.678587, -2.813661, -1.220141, 1.570796, 1.749976],accel_mss,speed_ms,0,blend_radius_m)
  movel([0.180554, -0.667081, -2.814913, -1.230395, 1.570796, 1.751350],accel_mss,speed_ms,0,blend_radius_m)
  movel([0.181390, -0.655935, -2.816072, -1.240382, 1.570796, 1.752186],accel_mss,speed_ms,0,blend_radius_m)
  movel([0.181508, -0.645334, -2.817127, -1.249928, 1.570796, 1.752305],accel_mss,speed_ms,0,blend_radius_m)
  movel([0.180716, -0.635477, -2.818066, -1.258846, 1.570796, 1.751512],accel_mss,speed_ms,0,blend_radius_m)
  movel([0.179492, -0.628855, -2.818676, -1.264858, 1.570796, 1.750288],accel_mss,speed_ms,0,blend_radius_m)
  movel([0.177674, -0.622575, -2.819237, -1.270577, 1.570796, 1.748470],accel_mss,speed_ms,0,blend_radius_m)
  movel([0.175212, -0.616814, -2.819738, -1.275836, 1.570796, 1.746008],accel_mss,speed_ms,0,blend_radius_m)
  movel([0.172054, -0.611754, -2.820168, -1.280467, 1.570796, 1.742851],accel_mss,speed_ms,0,blend_radius_m)
  movel([0.168163, -0.607565, -2.820516, -1.284308, 1.570796, 1.738959],accel_mss,speed_ms,0,blend_radius_m)
  movel([0.163499, -0.604415, -2.820773, -1.287201, 1.570796, 1.734295],accel_mss,speed_ms,0,blend_radius_m)
  movel([0.158021, -0.602490, -2.820928, -1.288971, 1.570796, 1.728817],accel_mss,speed_ms,0,blend_radius_m)
  movel([0.151716, -0.601943, -2.820972, -1.289473, 1.570796, 1.722513],accel_mss,speed_ms,0,blend_radius_m)
  movel([0.148431, -0.602267, -2.820946, -1.289176, 1.570796, 1.719227],accel_mss,speed_ms,0,blend_radius_m)
  movel([0.144882, -0.603048, -2.820884, -1.288457, 1.570796, 1.715678],accel_mss,speed_ms,0,blend_radius_m)
  movel([0.141095, -0.604309, -2.820782, -1.287298, 1.570796, 1.711892],accel_mss,speed_ms,0,blend_radius_m)
  movel([0.137112, -0.606061, -2.820639, -1.285689, 1.570796, 1.707908],accel_mss,speed_ms,0,blend_radius_m)
  movel([0.132975, -0.608300, -2.820455, -1.283634, 1.570796, 1.703772],accel_mss,speed_ms,0,blend_radius_m)
  movel([0.128708, -0.611053, -2.820227, -1.281110, 1.570796, 1.699505],accel_mss,speed_ms,0,blend_radius_m)
  movel([0.124362, -0.614309, -2.819952, -1.278128, 1.570796, 1.695159],accel_mss,speed_ms,0,blend_radius_m)
  movel([0.119974, -0.618083, -2.819629, -1.274677, 1.570796, 1.690770],accel_mss,speed_ms,0,blend_radius_m)
  speed_ms = 0.005
  movel([0.119974, -0.612246, -2.812827, -1.287316, 1.570796, 1.690770],accel_mss,speed_ms,0,blend_radius_m)
  speed_ms = 0.040
  movel([0.105668, -0.599555, -2.813887, -1.298947, 1.570796, 1.676464],accel_mss,speed_ms,0,blend_radius_m)
  speed_ms = 0.005
  movel([0.105668, -0.605180, -2.820711, -1.286498, 1.570796, 1.676464],accel_mss,speed_ms,0,blend_radius_m)
  speed_ms = 0.025
  movel([0.105208, -0.602800, -2.820903, -1.288686, 1.570796, 1.676004],accel_mss,speed_ms,0,blend_radius_m)
  movel([0.105101, -0.600110, -2.821118, -1.291161, 1.570796, 1.675897],accel_mss,speed_ms,0,blend_radius_m)
  movel([0.105749, -0.594005, -2.821596, -1.296788, 1.570796, 1.676545],accel_mss,speed_ms,0,blend_radius_m)
  movel([0.107230, -0.587216, -2.822110, -1.303063, 1.570796, 1.678026],accel_mss,speed_ms,0,blend_radius_m)
  movel([0.109136, -0.580136, -2.822627, -1.309626, 1.570796, 1.679932],accel_mss,speed_ms,0,blend_radius_m)
  speed_ms = 0.005
  movel([0.109136, -0.574935, -2.815764, -1.321690, 1.570796, 1.679932],accel_mss,speed_ms,0,blend_radius_m)
  speed_ms = 0.040
  movel([0.118580, -0.571553, -2.816004, -1.324833, 1.570796, 1.689376],accel_mss,speed_ms,0,blend_radius_m)
  speed_ms = 0.005
  movel([0.118580, -0.576694, -2.822872, -1.312823, 1.570796, 1.689376],accel_mss,speed_ms,0,blend_radius_m)
  speed_ms = 0.025
  movel([0.117402, -0.575267, -2.822972, -1.314150, 1.570796, 1.688198],accel_mss,speed_ms,0,blend_radius_m)
  movel([0.116582, -0.573518, -2.823093, -1.315777, 1.570796, 1.687379],accel_mss,speed_ms,0,blend_radius_m)
  movel([0.115918, -0.569140, -2.823393, -1.319856, 1.570796, 1.686715],accel_mss,speed_ms,0,blend_radius_m)
  movel([0.116427, -0.563751, -2.823752, -1.324886, 1.570796, 1.687223],accel_mss,speed_ms,0,blend_radius_m)
  movel([0.117944, -0.557530, -2.824152, -1.330706, 1.570796, 1.688741],accel_mss,speed_ms,0,blend_radius_m)
  movel([0.120304, -0.550672, -2.824578, -1.337139, 1.570796, 1.691100],accel_mss,speed_ms,0,blend_radius_m)
  movel([0.123332, -0.543377, -2.825011, -1.344000, 1.570796, 1.694129],accel_mss,speed_ms,0,blend_radius_m)
  movel([0.126853, -0.535849, -2.825438, -1.351102, 1.570796, 1.697649],accel_mss,speed_ms,0,blend_radius_m)
  movel([0.130680, -0.528304, -2.825846, -1.358240, 1.570796, 1.701476],accel_mss,speed_ms,0,blend_radius_m)
  speed_ms = 0.005
  movel([0.130680, -0.524028, -2.818917, -1.369444, 1.570796, 1.701476],accel_mss,speed_ms,0,blend_radius_m)
  speed_ms = 0.040
  movel([0.181260, -0.453275, -2.821737, -1.437377, 1.570796, 1.752057],accel_mss,speed_ms,0,blend_radius_m)
  speed_ms = 0.005
  movel([0.181260, -0.456170, -2.828726, -1.427493, 1.570796, 1.752057],accel_mss,speed_ms,0,blend_radius_m)
  speed_ms = 0.025
  movel([0.176078, -0.462124, -2.828557, -1.421708, 1.570796, 1.746874],accel_mss,speed_ms,0,blend_radius_m)
  movel([0.170926, -0.468393, -2.828365, -1.415631, 1.570796, 1.741722],accel_mss,speed_ms,0,blend_radius_m)
  movel([0.165890, -0.474874, -2.828153, -1.409362, 1.570796, 1.736686],accel_mss,speed_ms,0,blend_radius_m)
  movel([0.161028, -0.481494, -2.827921, -1.402974, 1.570796, 1.731824],accel_mss,speed_ms,0,blend_radius_m)
  movel([0.156423, -0.488161, -2.827672, -1.396555, 1.570796, 1.727219],accel_mss,speed_ms,0,blend_radius_m)
  movel([0.152136, -0.494789, -2.827410, -1.390190, 1.570796, 1.722932],accel_mss,speed_ms,0,blend_radius_m)
  movel([0.148234, -0.501305, -2.827137, -1.383947, 1.570796, 1.719030],accel_mss,speed_ms,0,blend_radius_m)
  movel([0.144778, -0.507634, -2.826857, -1.377898, 1.570796, 1.715575],accel_mss,speed_ms,0,blend_radius_m)
  movel([0.141828, -0.513689, -2.826577, -1.372124, 1.570796, 1.712624],accel_mss,speed_ms,0,blend_radius_m)
  movel([0.139435, -0.519412, -2.826300, -1.366678, 1.570796, 1.710232],accel_mss,speed_ms,0,blend_radius_m)
  movel([0.137657, -0.524728, -2.826032, -1.361629, 1.570796, 1.708453],accel_mss,speed_ms,0,blend_radius_m)
  movel([0.136544, -0.529571, -2.825779, -1.357039, 1.570796, 1.707340],accel_mss,speed_ms,0,blend_radius_m)
  movel([0.136155, -0.533872, -2.825547, -1.352970, 1.570796, 1.706952],accel_mss,speed_ms,0,blend_radius_m)
  movel([0.136543, -0.537565, -2.825343, -1.349481, 1.570796, 1.707339],accel_mss,speed_ms,0,blend_radius_m)
  movel([0.137752, -0.540595, -2.825171, -1.346623, 1.570796, 1.708548],accel_mss,speed_ms,0,blend_radius_m)
  movel([0.139843, -0.542894, -2.825039, -1.344456, 1.570796, 1.710639],accel_mss,speed_ms,0,blend_radius_m)
  speed_ms = 0.005
  movel([0.139843, -0.538352, -2.818127, -1.355910, 1.570796, 1.710639],accel_mss,speed_ms,0,blend_radius_m)
  speed_ms = 0.040
  movel([0.162855, -0.512881, -2.819479, -1.380028, 1.570796, 1.733652],accel_mss,speed_ms,0,blend_radius_m)
  speed_ms = 0.005
  movel([0.162855, -0.516946, -2.826420, -1.369023, 1.570796, 1.733652],accel_mss,speed_ms,0,blend_radius_m)
  speed_ms = 0.025
  movel([0.162384, -0.514031, -2.826561, -1.371797, 1.570796, 1.733180],accel_mss,speed_ms,0,blend_radius_m)
  movel([0.162288, -0.510755, -2.826714, -1.374920, 1.570796, 1.733084],accel_mss,speed_ms,0,blend_radius_m)
  movel([0.162565, -0.507153, -2.826879, -1.378357, 1.570796, 1.733362],accel_mss,speed_ms,0,blend_radius_m)
  movel([0.163216, -0.503245, -2.827053, -1.382092, 1.570796, 1.734012],accel_mss,speed_ms,0,blend_radius_m)
  movel([0.164233, -0.499067, -2.827232, -1.386090, 1.570796, 1.735029],accel_mss,speed_ms,0,blend_radius_m)
  movel([0.165623, -0.494639, -2.827416, -1.390334, 1.570796, 1.736419],accel_mss,speed_ms,0,blend_radius_m)
  movel([0.167387, -0.489981, -2.827602, -1.394806, 1.570796, 1.738183],accel_mss,speed_ms,0,blend_radius_m)
  movel([0.169516, -0.485137, -2.827787, -1.399465, 1.570796, 1.740313],accel_mss,speed_ms,0,blend_radius_m)
  movel([0.172012, -0.480127, -2.827970, -1.404292, 1.570796, 1.742809],accel_mss,speed_ms,0,blend_radius_m)
  movel([0.174881, -0.474973, -2.828149, -1.409266, 1.570796, 1.745678],accel_mss,speed_ms,0,blend_radius_m)
  movel([0.178106, -0.469729, -2.828322, -1.414338, 1.570796, 1.748902],accel_mss,speed_ms,0,blend_radius_m)
  movel([0.181701, -0.464399, -2.828489, -1.419501, 1.570796, 1.752497],accel_mss,speed_ms,0,blend_radius_m)
  movel([0.185655, -0.459027, -2.828646, -1.424716, 1.570796, 1.756451],accel_mss,speed_ms,0,blend_radius_m)
  movel([0.189965, -0.453644, -2.828794, -1.429951, 1.570796, 1.760761],accel_mss,speed_ms,0,blend_radius_m)
  movel([0.194624, -0.448291, -2.828932, -1.435166, 1.570796, 1.765421],accel_mss,speed_ms,0,blend_radius_m)
  movel([0.199621, -0.443002, -2.829058, -1.440329, 1.570796, 1.770417],accel_mss,speed_ms,0,blend_radius_m)
  movel([0.204634, -0.438137, -2.829166, -1.445086, 1.570796, 1.775430],accel_mss,speed_ms,0,blend_radius_m)
  movel([0.209620, -0.433721, -2.829257, -1.449411, 1.570796, 1.780416],accel_mss,speed_ms,0,blend_radius_m)
  movel([0.214539, -0.429759, -2.829333, -1.453297, 1.570796, 1.785336],accel_mss,speed_ms,0,blend_radius_m)
  movel([0.219373, -0.426252, -2.829395, -1.456741, 1.570796, 1.790170],accel_mss,speed_ms,0,blend_radius_m)
  movel([0.224084, -0.423203, -2.829447, -1.459739, 1.570796, 1.794880],accel_mss,speed_ms,0,blend_radius_m)
  movel([0.228628, -0.420629, -2.829488, -1.462273, 1.570796, 1.799425],accel_mss,speed_ms,0,blend_radius_m)
  movel([0.232995, -0.418506, -2.829520, -1.464364, 1.570796, 1.803792],accel_mss,speed_ms,0,blend_radius_m)
  movel([0.237129, -0.416859, -2.829543, -1.465986, 1.570796, 1.807925],accel_mss,speed_ms,0,blend_radius_m)
  movel([0.241016, -0.415678, -2.829560, -1.467151, 1.570796, 1.811812],accel_mss,speed_ms,0,blend_radius_m)
  movel([0.247935, -0.414689, -2.829573, -1.468127, 1.570796, 1.818732],accel_mss,speed_ms,0,blend_radius_m)
  movel([0.250900, -0.414885, -2.829571, -1.467933, 1.570796, 1.821697],accel_mss,speed_ms,0,blend_radius_m)
  movel([0.255753, -0.416602, -2.829547, -1.466240, 1.570796, 1.826549],accel_mss,speed_ms,0,blend_radius_m)
  movel([0.257590, -0.418106, -2.829525, -1.464758, 1.570796, 1.828387],accel_mss,speed_ms,0,blend_radius_m)
  movel([0.259001, -0.420034, -2.829497, -1.462858, 1.570796, 1.829798],accel_mss,speed_ms,0,blend_radius_m)
  speed_ms = 0.005
  movel([0.259001, -0.417864, -2.822491, -1.472034, 1.570796, 1.829798],accel_mss,speed_ms,0,blend_radius_m)
  speed_ms = 0.040
  movel([0.274724, -0.430831, -2.822265, -1.459293, 1.570796, 1.845520],accel_mss,speed_ms,0,blend_radius_m)
  speed_ms = 0.005
  movel([0.274724, -0.433269, -2.829266, -1.449855, 1.570796, 1.845520],accel_mss,speed_ms,0,blend_radius_m)
  speed_ms = 0.025
  movel([0.272812, -0.430079, -2.829327, -1.452983, 1.570796, 1.843609],accel_mss,speed_ms,0,blend_radius_m)
  movel([0.269936, -0.428053, -2.829364, -1.454972, 1.570796, 1.840732],accel_mss,speed_ms,0,blend_radius_m)
  movel([0.266170, -0.427187, -2.829379, -1.455823, 1.570796, 1.836967],accel_mss,speed_ms,0,blend_radius_m)
  movel([0.261578, -0.427480, -2.829374, -1.455536, 1.570796, 1.832374],accel_mss,speed_ms,0,blend_radius_m)
  movel([0.256264, -0.428903, -2.829348, -1.454138, 1.570796, 1.827060],accel_mss,speed_ms,0,blend_radius_m)
  movel([0.250302, -0.431450, -2.829301, -1.451639, 1.570796, 1.821099],accel_mss,speed_ms,0,blend_radius_m)
  movel([0.243802, -0.435085, -2.829229, -1.448075, 1.570796, 1.814599],accel_mss,speed_ms,0,blend_radius_m)
  movel([0.236850, -0.439782, -2.829130, -1.443477, 1.570796, 1.807647],accel_mss,speed_ms,0,blend_radius_m)
  movel([0.229570, -0.445491, -2.829000, -1.437898, 1.570796, 1.800366],accel_mss,speed_ms,0,blend_radius_m)
  movel([0.222137, -0.452098, -2.828835, -1.431456, 1.570796, 1.792933],accel_mss,speed_ms,0,blend_radius_m)
  movel([0.214847, -0.459360, -2.828637, -1.424392, 1.570796, 1.785644],accel_mss,speed_ms,0,blend_radius_m)
  movel([0.208004, -0.467046, -2.828407, -1.416936, 1.570796, 1.778801],accel_mss,speed_ms,0,blend_radius_m)
  movel([0.201871, -0.474943, -2.828150, -1.409295, 1.570796, 1.772667],accel_mss,speed_ms,0,blend_radius_m)
  movel([0.199162, -0.478898, -2.828014, -1.405477, 1.570796, 1.769958],accel_mss,speed_ms,0,blend_radius_m)
  movel([0.196726, -0.482824, -2.827873, -1.401692, 1.570796, 1.767523],accel_mss,speed_ms,0,blend_radius_m)
  movel([0.194595, -0.486701, -2.827728, -1.397960, 1.570796, 1.765391],accel_mss,speed_ms,0,blend_radius_m)
  movel([0.192805, -0.490505, -2.827581, -1.394302, 1.570796, 1.763601],accel_mss,speed_ms,0,blend_radius_m)
  movel([0.191376, -0.494210, -2.827433, -1.390745, 1.570796, 1.762173],accel_mss,speed_ms,0,blend_radius_m)
  movel([0.190353, -0.497782, -2.827286, -1.387320, 1.570796, 1.761149],accel_mss,speed_ms,0,blend_radius_m)
  speed_ms = 0.005
  movel([0.190353, -0.494079, -2.820327, -1.397982, 1.570796, 1.761149],accel_mss,speed_ms,0,blend_radius_m)
  speed_ms = 0.040
  movel([0.225557, -0.482976, -2.820769, -1.408644, 1.570796, 1.796354],accel_mss,speed_ms,0,blend_radius_m)
  speed_ms = 0.005
  movel([0.225557, -0.486462, -2.827737, -1.398189, 1.570796, 1.796354],accel_mss,speed_ms,0,blend_radius_m)
  speed_ms = 0.025
  movel([0.230532, -0.480919, -2.827942, -1.403528, 1.570796, 1.801329],accel_mss,speed_ms,0,blend_radius_m)
  movel([0.235675, -0.475846, -2.828120, -1.408423, 1.570796, 1.806472],accel_mss,speed_ms,0,blend_radius_m)
  movel([0.240904, -0.471270, -2.828273, -1.412847, 1.570796, 1.811700],accel_mss,speed_ms,0,blend_radius_m)
  movel([0.246113, -0.467241, -2.828401, -1.416747, 1.570796, 1.816909],accel_mss,speed_ms,0,blend_radius_m)
  movel([0.251210, -0.463791, -2.828507, -1.420091, 1.570796, 1.822007],accel_mss,speed_ms,0,blend_radius_m)
  movel([0.256093, -0.460955, -2.828591, -1.422843, 1.570796, 1.826889],accel_mss,speed_ms,0,blend_radius_m)
  movel([0.260676, -0.458762, -2.828654, -1.424974, 1.570796, 1.831472],accel_mss,speed_ms,0,blend_radius_m)
  movel([0.264851, -0.457246, -2.828696, -1.426447, 1.570796, 1.835647],accel_mss,speed_ms,0,blend_radius_m)
  movel([0.269216, -0.456489, -2.828717, -1.427183, 1.570796, 1.840012],accel_mss,speed_ms,0,blend_radius_m)
  movel([0.272323, -0.457089, -2.828701, -1.426599, 1.570796, 1.843120],accel_mss,speed_ms,0,blend_radius_m)
  movel([0.274310, -0.458896, -2.828650, -1.424843, 1.570796, 1.845106],accel_mss,speed_ms,0,blend_radius_m)
  movel([0.275291, -0.461777, -2.828567, -1.422045, 1.570796, 1.846087],accel_mss,speed_ms,0,blend_radius_m)
  movel([0.275404, -0.465568, -2.828453, -1.418368, 1.570796, 1.846201],accel_mss,speed_ms,0,blend_radius_m)
  movel([0.274782, -0.470132, -2.828309, -1.413947, 1.570796, 1.845579],accel_mss,speed_ms,0,blend_radius_m)
  movel([0.273555, -0.475317, -2.828138, -1.408934, 1.570796, 1.844351],accel_mss,speed_ms,0,blend_radius_m)
  movel([0.271863, -0.480972, -2.827940, -1.403477, 1.570796, 1.842660],accel_mss,speed_ms,0,blend_radius_m)
  speed_ms = 0.005
  movel([0.271863, -0.477592, -2.820967, -1.413830, 1.570796, 1.842660],accel_mss,speed_ms,0,blend_radius_m)
  speed_ms = 0.040
  movel([0.237934, -0.497934, -2.820164, -1.394291, 1.570796, 1.808730],accel_mss,speed_ms,0,blend_radius_m)
  speed_ms = 0.005
  movel([0.237934, -0.501712, -2.827119, -1.383558, 1.570796, 1.808730],accel_mss,speed_ms,0,blend_radius_m)
  speed_ms = 0.025
  movel([0.242451, -0.499306, -2.827222, -1.385861, 1.570796, 1.813247],accel_mss,speed_ms,0,blend_radius_m)
  movel([0.246530, -0.497618, -2.827293, -1.387478, 1.570796, 1.817326],accel_mss,speed_ms,0,blend_radius_m)
  movel([0.250167, -0.496633, -2.827334, -1.388422, 1.570796, 1.820964],accel_mss,speed_ms,0,blend_radius_m)
  movel([0.253371, -0.496299, -2.827348, -1.388742, 1.570796, 1.824168],accel_mss,speed_ms,0,blend_radius_m)
  movel([0.256145, -0.496592, -2.827336, -1.388461, 1.570796, 1.826941],accel_mss,speed_ms,0,blend_radius_m)
  movel([0.258492, -0.497468, -2.827299, -1.387621, 1.570796, 1.829288],accel_mss,speed_ms,0,blend_radius_m)
  movel([0.260428, -0.498888, -2.827240, -1.386261, 1.570796, 1.831224],accel_mss,speed_ms,0,blend_radius_m)
  movel([0.261949, -0.500825, -2.827158, -1.384407, 1.570796, 1.832745],accel_mss,speed_ms,0,blend_radius_m)
  movel([0.263082, -0.503224, -2.827054, -1.382112, 1.570796, 1.833878],accel_mss,speed_ms,0,blend_radius_m)
  movel([0.263834, -0.506045, -2.826929, -1.379415, 1.570796, 1.834630],accel_mss,speed_ms,0,blend_radius_m)
  movel([0.264212, -0.509256, -2.826784, -1.376350, 1.570796, 1.835008],accel_mss,speed_ms,0,blend_radius_m)
  movel([0.264237, -0.512805, -2.826619, -1.372966, 1.570796, 1.835033],accel_mss,speed_ms,0,blend_radius_m)
  movel([0.263917, -0.516659, -2.826434, -1.369296, 1.570796, 1.834713],accel_mss,speed_ms,0,blend_radius_m)
  movel([0.262305, -0.525101, -2.826012, -1.361276, 1.570796, 1.833101],accel_mss,speed_ms,0,blend_radius_m)
  movel([0.261033, -0.529618, -2.825776, -1.356995, 1.570796, 1.831830],accel_mss,speed_ms,0,blend_radius_m)
  movel([0.260911, -0.528484, -2.825836, -1.358069, 1.570796, 1.831708],accel_mss,speed_ms,0,blend_radius_m)
  speed_ms = 0.005
  movel([0.260911, -0.524205, -2.818907, -1.369276, 1.570796, 1.831708],accel_mss,speed_ms,0,blend_radius_m)
  speed_ms = 0.040
  movel([0.286425, -0.522747, -2.818984, -1.370659, 1.570796, 1.857221],accel_mss,speed_ms,0,blend_radius_m)
  speed_ms = 0.005
  movel([0.286425, -0.526998, -2.825914, -1.359477, 1.570796, 1.857221],accel_mss,speed_ms,0,blend_radius_m)
  speed_ms = 0.025
  movel([0.281721, -0.534373, -2.825520, -1.352496, 1.570796, 1.852517],accel_mss,speed_ms,0,blend_radius_m)
  movel([0.277579, -0.541642, -2.825112, -1.345636, 1.570796, 1.848375],accel_mss,speed_ms,0,blend_radius_m)
  movel([0.273882, -0.548783, -2.824692, -1.338914, 1.570796, 1.844679],accel_mss,speed_ms,0,blend_radius_m)
  movel([0.270506, -0.555784, -2.824262, -1.332342, 1.570796, 1.841302],accel_mss,speed_ms,0,blend_radius_m)
  movel([0.267119, -0.563333, -2.823779, -1.325277, 1.570796, 1.837915],accel_mss,speed_ms,0,blend_radius_m)
  movel([0.265729, -0.566940, -2.823541, -1.321908, 1.570796, 1.836525],accel_mss,speed_ms,0,blend_radius_m)
  movel([0.264664, -0.570356, -2.823310, -1.318722, 1.570796, 1.835460],accel_mss,speed_ms,0,blend_radius_m)
  movel([0.264005, -0.573513, -2.823094, -1.315782, 1.570796, 1.834801],accel_mss,speed_ms,0,blend_radius_m)
  movel([0.263849, -0.576274, -2.822901, -1.313214, 1.570796, 1.834645],accel_mss,speed_ms,0,blend_radius_m)
  movel([0.264284, -0.578464, -2.822746, -1.311178, 1.570796, 1.835080],accel_mss,speed_ms,0,blend_radius_m)
  movel([0.265378, -0.579943, -2.822641, -1.309805, 1.570796, 1.836174],accel_mss,speed_ms,0,blend_radius_m)
  movel([0.268144, -0.580963, -2.822567, -1.308858, 1.570796, 1.838940],accel_mss,speed_ms,0,blend_radius_m)
  movel([0.269503, -0.581492, -2.822529, -1.308368, 1.570796, 1.840299],accel_mss,speed_ms,0,blend_radius_m)
  movel([0.270510, -0.582456, -2.822459, -1.307473, 1.570796, 1.841306],accel_mss,speed_ms,0,blend_radius_m)
  movel([0.270926, -0.584415, -2.822317, -1.305657, 1.570796, 1.841723],accel_mss,speed_ms,0,blend_radius_m)
  movel([0.270622, -0.587231, -2.822109, -1.303049, 1.570796, 1.841419],accel_mss,speed_ms,0,blend_radius_m)
  movel([0.269763, -0.590672, -2.821850, -1.299866, 1.570796, 1.840560],accel_mss,speed_ms,0,blend_radius_m)
  movel([0.268504, -0.594506, -2.821557, -1.296326, 1.570796, 1.839300],accel_mss,speed_ms,0,blend_radius_m)
  movel([0.265395, -0.602462, -2.820931, -1.288997, 1.570796, 1.836191],accel_mss,speed_ms,0,blend_radius_m)
  movel([0.255783, -0.624793, -2.819041, -1.268555, 1.570796, 1.826579],accel_mss,speed_ms,0,blend_radius_m)
  movel([0.249309, -0.639979, -2.817642, -1.254767, 1.570796, 1.820106],accel_mss,speed_ms,0,blend_radius_m)
  movel([0.247618, -0.644499, -2.817208, -1.250682, 1.570796, 1.818415],accel_mss,speed_ms,0,blend_radius_m)
  movel([0.246095, -0.649195, -2.816748, -1.246446, 1.570796, 1.816891],accel_mss,speed_ms,0,blend_radius_m)
  movel([0.243703, -0.658696, -2.815790, -1.237903, 1.570796, 1.814500],accel_mss,speed_ms,0,blend_radius_m)
  movel([0.242917, -0.663297, -2.815312, -1.233780, 1.570796, 1.813713],accel_mss,speed_ms,0,blend_radius_m)
  movel([0.242456, -0.667660, -2.814851, -1.229878, 1.570796, 1.813252],accel_mss,speed_ms,0,blend_radius_m)
  movel([0.242353, -0.671688, -2.814418, -1.226282, 1.570796, 1.813149],accel_mss,speed_ms,0,blend_radius_m)
  movel([0.242645, -0.675290, -2.814025, -1.223074, 1.570796, 1.813442],accel_mss,speed_ms,0,blend_radius_m)
  movel([0.243374, -0.678355, -2.813687, -1.220348, 1.570796, 1.814170],accel_mss,speed_ms,0,blend_radius_m)
  movel([0.244568, -0.680806, -2.813413, -1.218170, 1.570796, 1.815364],accel_mss,speed_ms,0,blend_radius_m)
  movel([0.246276, -0.682531, -2.813219, -1.216639, 1.570796, 1.817072],accel_mss,speed_ms,0,blend_radius_m)
  movel([0.248533, -0.683440, -2.813116, -1.215833, 1.570796, 1.819329],accel_mss,speed_ms,0,blend_radius_m)
  movel([0.251378, -0.683435, -2.813117, -1.215838, 1.570796, 1.822174],accel_mss,speed_ms,0,blend_radius_m)
  movel([0.254864, -0.682409, -2.813233, -1.216747, 1.570796, 1.825661],accel_mss,speed_ms,0,blend_radius_m)
  movel([0.259038, -0.680262, -2.813474, -1.218653, 1.570796, 1.829835],accel_mss,speed_ms,0,blend_radius_m)
  movel([0.263958, -0.676881, -2.813850, -1.221658, 1.570796, 1.834754],accel_mss,speed_ms,0,blend_radius_m)
  movel([0.267886, -0.673675, -2.814202, -1.224512, 1.570796, 1.838682],accel_mss,speed_ms,0,blend_radius_m)
  movel([0.271783, -0.670109, -2.814589, -1.227692, 1.570796, 1.842579],accel_mss,speed_ms,0,blend_radius_m)
  movel([0.275661, -0.666230, -2.815003, -1.231156, 1.570796, 1.846457],accel_mss,speed_ms,0,blend_radius_m)
  movel([0.279521, -0.662100, -2.815437, -1.234852, 1.570796, 1.850318],accel_mss,speed_ms,0,blend_radius_m)
  movel([0.287206, -0.653327, -2.816336, -1.242726, 1.570796, 1.858002],accel_mss,speed_ms,0,blend_radius_m)
  movel([0.294865, -0.644277, -2.817229, -1.250883, 1.570796, 1.865661],accel_mss,speed_ms,0,blend_radius_m)
  movel([0.302757, -0.635238, -2.818089, -1.259062, 1.570796, 1.873553],accel_mss,speed_ms,0,blend_radius_m)
  movel([0.306845, -0.630834, -2.818495, -1.263060, 1.570796, 1.877642],accel_mss,speed_ms,0,blend_radius_m)
  movel([0.310988, -0.626636, -2.818876, -1.266877, 1.570796, 1.881784],accel_mss,speed_ms,0,blend_radius_m)
  movel([0.315153, -0.622729, -2.819224, -1.270437, 1.570796, 1.885950],accel_mss,speed_ms,0,blend_radius_m)
  movel([0.319307, -0.619218, -2.819531, -1.273640, 1.570796, 1.890104],accel_mss,speed_ms,0,blend_radius_m)
  movel([0.323408, -0.616199, -2.819791, -1.276398, 1.570796, 1.894204],accel_mss,speed_ms,0,blend_radius_m)
  movel([0.327424, -0.613774, -2.819998, -1.278617, 1.570796, 1.898220],accel_mss,speed_ms,0,blend_radius_m)
  movel([0.335704, -0.610053, -2.820310, -1.282025, 1.570796, 1.906501],accel_mss,speed_ms,0,blend_radius_m)
  movel([0.338553, -0.608565, -2.820434, -1.283391, 1.570796, 1.909349],accel_mss,speed_ms,0,blend_radius_m)
  movel([0.341622, -0.606491, -2.820604, -1.285294, 1.570796, 1.912418],accel_mss,speed_ms,0,blend_radius_m)
  movel([0.344775, -0.603786, -2.820824, -1.287779, 1.570796, 1.915572],accel_mss,speed_ms,0,blend_radius_m)
  movel([0.347727, -0.600584, -2.821081, -1.290724, 1.570796, 1.918524],accel_mss,speed_ms,0,blend_radius_m)
  movel([0.349043, -0.598830, -2.821220, -1.292340, 1.570796, 1.919839],accel_mss,speed_ms,0,blend_radius_m)
  movel([0.350203, -0.596999, -2.821363, -1.294027, 1.570796, 1.920999],accel_mss,speed_ms,0,blend_radius_m)
  speed_ms = 0.005
  movel([0.350203, -0.591510, -2.814526, -1.306353, 1.570796, 1.920999],accel_mss,speed_ms,0,blend_radius_m)
  speed_ms = 0.040
  movel([0.368105, -0.558133, -2.816912, -1.337344, 1.570796, 1.938901],accel_mss,speed_ms,0,blend_radius_m)
  speed_ms = 0.005
  movel([0.368105, -0.563036, -2.823798, -1.325555, 1.570796, 1.938901],accel_mss,speed_ms,0,blend_radius_m)
  speed_ms = 0.025
  movel([0.368968, -0.563108, -2.823794, -1.325487, 1.570796, 1.939765],accel_mss,speed_ms,0,blend_radius_m)
  movel([0.368864, -0.564341, -2.823713, -1.324335, 1.570796, 1.939660],accel_mss,speed_ms,0,blend_radius_m)
  movel([0.368010, -0.566157, -2.823593, -1.322639, 1.570796, 1.938806],accel_mss,speed_ms,0,blend_radius_m)
  movel([0.366650, -0.567975, -2.823471, -1.320942, 1.570796, 1.937447],accel_mss,speed_ms,0,blend_radius_m)
  movel([0.365112, -0.569397, -2.823375, -1.319616, 1.570796, 1.935908],accel_mss,speed_ms,0,blend_radius_m)
  movel([0.363581, -0.570507, -2.823300, -1.318582, 1.570796, 1.934377],accel_mss,speed_ms,0,blend_radius_m)
  movel([0.360546, -0.572401, -2.823170, -1.316818, 1.570796, 1.931342],accel_mss,speed_ms,0,blend_radius_m)
  movel([0.358317, -0.574025, -2.823058, -1.315306, 1.570796, 1.929113],accel_mss,speed_ms,0,blend_radius_m)
  movel([0.356086, -0.575943, -2.822924, -1.313521, 1.570796, 1.926882],accel_mss,speed_ms,0,blend_radius_m)
  movel([0.351647, -0.580448, -2.822605, -1.309337, 1.570796, 1.922443],accel_mss,speed_ms,0,blend_radius_m)
  movel([0.347317, -0.585512, -2.822236, -1.304641, 1.570796, 1.918113],accel_mss,speed_ms,0,blend_radius_m)
  movel([0.343182, -0.590709, -2.821847, -1.299833, 1.570796, 1.913979],accel_mss,speed_ms,0,blend_radius_m)
  movel([0.342235, -0.591999, -2.821749, -1.298640, 1.570796, 1.913032],accel_mss,speed_ms,0,blend_radius_m)
  movel([0.341615, -0.593220, -2.821656, -1.297513, 1.570796, 1.912411],accel_mss,speed_ms,0,blend_radius_m)
  movel([0.341723, -0.594101, -2.821588, -1.296700, 1.570796, 1.912520],accel_mss,speed_ms,0,blend_radius_m)
  movel([0.342462, -0.594340, -2.821570, -1.296479, 1.570796, 1.913258],accel_mss,speed_ms,0,blend_radius_m)
  movel([0.344503, -0.594228, -2.821578, -1.296583, 1.570796, 1.915299],accel_mss,speed_ms,0,blend_radius_m)
  movel([0.346807, -0.593628, -2.821625, -1.297137, 1.570796, 1.917604],accel_mss,speed_ms,0,blend_radius_m)
  movel([0.349334, -0.592575, -2.821705, -1.298108, 1.570796, 1.920130],accel_mss,speed_ms,0,blend_radius_m)
  movel([0.352037, -0.591085, -2.821819, -1.299485, 1.570796, 1.922833],accel_mss,speed_ms,0,blend_radius_m)
  movel([0.354856, -0.589207, -2.821961, -1.301222, 1.570796, 1.925652],accel_mss,speed_ms,0,blend_radius_m)
  movel([0.357752, -0.586950, -2.822129, -1.303309, 1.570796, 1.928549],accel_mss,speed_ms,0,blend_radius_m)
  movel([0.360668, -0.584358, -2.822321, -1.305710, 1.570796, 1.931464],accel_mss,speed_ms,0,blend_radius_m)
  movel([0.363561, -0.581446, -2.822533, -1.308410, 1.570796, 1.934358],accel_mss,speed_ms,0,blend_radius_m)
  movel([0.362934, -0.583249, -2.822402, -1.306738, 1.570796, 1.933731],accel_mss,speed_ms,0,blend_radius_m)
  movel([0.363038, -0.584522, -2.822309, -1.305559, 1.570796, 1.933835],accel_mss,speed_ms,0,blend_radius_m)
  movel([0.363749, -0.585192, -2.822259, -1.304938, 1.570796, 1.934545],accel_mss,speed_ms,0,blend_radius_m)
  movel([0.364933, -0.585192, -2.822259, -1.304938, 1.570796, 1.935729],accel_mss,speed_ms,0,blend_radius_m)
  movel([0.366423, -0.584574, -2.822305, -1.305510, 1.570796, 1.937220],accel_mss,speed_ms,0,blend_radius_m)
  movel([0.368082, -0.583530, -2.822381, -1.306477, 1.570796, 1.938878],accel_mss,speed_ms,0,blend_radius_m)
  movel([0.371589, -0.580648, -2.822590, -1.309151, 1.570796, 1.942385],accel_mss,speed_ms,0,blend_radius_m)
  movel([0.376077, -0.576275, -2.822901, -1.313213, 1.570796, 1.946874],accel_mss,speed_ms,0,blend_radius_m)
  movel([0.380438, -0.571407, -2.823239, -1.317743, 1.570796, 1.951234],accel_mss,speed_ms,0,blend_radius_m)
  movel([0.384550, -0.566191, -2.823591, -1.322607, 1.570796, 1.955347],accel_mss,speed_ms,0,blend_radius_m)
  movel([0.388290, -0.560770, -2.823946, -1.327674, 1.570796, 1.959086],accel_mss,speed_ms,0,blend_radius_m)
  movel([0.389384, -0.558928, -2.824064, -1.329398, 1.570796, 1.960180],accel_mss,speed_ms,0,blend_radius_m)
  movel([0.389964, -0.557329, -2.824165, -1.330895, 1.570796, 1.960761],accel_mss,speed_ms,0,blend_radius_m)
  movel([0.389788, -0.556499, -2.824218, -1.331672, 1.570796, 1.960584],accel_mss,speed_ms,0,blend_radius_m)
  movel([0.389203, -0.556103, -2.824242, -1.332044, 1.570796, 1.959999],accel_mss,speed_ms,0,blend_radius_m)
  movel([0.386676, -0.555568, -2.824276, -1.332545, 1.570796, 1.957472],accel_mss,speed_ms,0,blend_radius_m)
  movel([0.381451, -0.555387, -2.824287, -1.332715, 1.570796, 1.952247],accel_mss,speed_ms,0,blend_radius_m)
  movel([0.379326, -0.554280, -2.824356, -1.333753, 1.570796, 1.950122],accel_mss,speed_ms,0,blend_radius_m)
  movel([0.384469, -0.548245, -2.824724, -1.339420, 1.570796, 1.955266],accel_mss,speed_ms,0,blend_radius_m)
  movel([0.387180, -0.545539, -2.824885, -1.341965, 1.570796, 1.957976],accel_mss,speed_ms,0,blend_radius_m)
  movel([0.389910, -0.543219, -2.825020, -1.344149, 1.570796, 1.960706],accel_mss,speed_ms,0,blend_radius_m)
  movel([0.391735, -0.541964, -2.825093, -1.345332, 1.570796, 1.962531],accel_mss,speed_ms,0,blend_radius_m)
  movel([0.393582, -0.540946, -2.825151, -1.346292, 1.570796, 1.964378],accel_mss,speed_ms,0,blend_radius_m)
  movel([0.396744, -0.539878, -2.825212, -1.347299, 1.570796, 1.967540],accel_mss,speed_ms,0,blend_radius_m)
  movel([0.398201, -0.540302, -2.825188, -1.346898, 1.570796, 1.968997],accel_mss,speed_ms,0,blend_radius_m)
  movel([0.398494, -0.541030, -2.825147, -1.346212, 1.570796, 1.969291],accel_mss,speed_ms,0,blend_radius_m)
  movel([0.398393, -0.542125, -2.825084, -1.345180, 1.570796, 1.969189],accel_mss,speed_ms,0,blend_radius_m)
  movel([0.397663, -0.543938, -2.824979, -1.343472, 1.570796, 1.968460],accel_mss,speed_ms,0,blend_radius_m)
  movel([0.396447, -0.545918, -2.824862, -1.341608, 1.570796, 1.967243],accel_mss,speed_ms,0,blend_radius_m)
  movel([0.393297, -0.549885, -2.824626, -1.337879, 1.570796, 1.964093],accel_mss,speed_ms,0,blend_radius_m)
  speed_ms = 0.005
  movel([0.393297, -0.545216, -2.817722, -1.349451, 1.570796, 1.964093],accel_mss,speed_ms,0,blend_radius_m)
  speed_ms = 0.040
  movel([0.440057, -0.418094, -2.822487, -1.471807, 1.570796, 2.010854],accel_mss,speed_ms,0,blend_radius_m)
  speed_ms = 0.005
  movel([0.440057, -0.420270, -2.829493, -1.462626, 1.570796, 2.010854],accel_mss,speed_ms,0,blend_radius_m)
  speed_ms = 0.025
  movel([0.442441, -0.418079, -2.829526, -1.464784, 1.570796, 2.013238],accel_mss,speed_ms,0,blend_radius_m)
  movel([0.444761, -0.416261, -2.829552, -1.466576, 1.570796, 2.015558],accel_mss,speed_ms,0,blend_radius_m)
  movel([0.446970, -0.414822, -2.829572, -1.467995, 1.570796, 2.017767],accel_mss,speed_ms,0,blend_radius_m)
  movel([0.450910, -0.413094, -2.829594, -1.469701, 1.570796, 2.021706],accel_mss,speed_ms,0,blend_radius_m)
  movel([0.452557, -0.412808, -2.829598, -1.469983, 1.570796, 2.023353],accel_mss,speed_ms,0,blend_radius_m)
  movel([0.455003, -0.413405, -2.829590, -1.469393, 1.570796, 2.025800],accel_mss,speed_ms,0,blend_radius_m)
  movel([0.456272, -0.415371, -2.829564, -1.467454, 1.570796, 2.027069],accel_mss,speed_ms,0,blend_radius_m)
  movel([0.456587, -0.418332, -2.829522, -1.464535, 1.570796, 2.027383],accel_mss,speed_ms,0,blend_radius_m)
  movel([0.456142, -0.422020, -2.829466, -1.460904, 1.570796, 2.026938],accel_mss,speed_ms,0,blend_radius_m)
  movel([0.455131, -0.426170, -2.829397, -1.456822, 1.570796, 2.025928],accel_mss,speed_ms,0,blend_radius_m)
  movel([0.452847, -0.432981, -2.829271, -1.450137, 1.570796, 2.023643],accel_mss,speed_ms,0,blend_radius_m)
  movel([0.449787, -0.440277, -2.829119, -1.442993, 1.570796, 2.020584],accel_mss,speed_ms,0,blend_radius_m)
  movel([0.446023, -0.447926, -2.828941, -1.435523, 1.570796, 2.016820],accel_mss,speed_ms,0,blend_radius_m)
  movel([0.437383, -0.463249, -2.828523, -1.420617, 1.570796, 2.008179],accel_mss,speed_ms,0,blend_radius_m)
  movel([0.435923, -0.466566, -2.828422, -1.417401, 1.570796, 2.006720],accel_mss,speed_ms,0,blend_radius_m)
  movel([0.435426, -0.469203, -2.828339, -1.414847, 1.570796, 2.006222],accel_mss,speed_ms,0,blend_radius_m)
  movel([0.435982, -0.470660, -2.828292, -1.413436, 1.570796, 2.006778],accel_mss,speed_ms,0,blend_radius_m)
  movel([0.437126, -0.471482, -2.828266, -1.412642, 1.570796, 2.007923],accel_mss,speed_ms,0,blend_radius_m)
  movel([0.438392, -0.472184, -2.828243, -1.411963, 1.570796, 2.009189],accel_mss,speed_ms,0,blend_radius_m)
  movel([0.439295, -0.473292, -2.828206, -1.410891, 1.570796, 2.010091],accel_mss,speed_ms,0,blend_radius_m)
  movel([0.439487, -0.474920, -2.828151, -1.409317, 1.570796, 2.010284],accel_mss,speed_ms,0,blend_radius_m)
  movel([0.439143, -0.477033, -2.828079, -1.407278, 1.570796, 2.009939],accel_mss,speed_ms,0,blend_radius_m)
  movel([0.437530, -0.481993, -2.827903, -1.402493, 1.570796, 2.008326],accel_mss,speed_ms,0,blend_radius_m)
  movel([0.434579, -0.489482, -2.827621, -1.395285, 1.570796, 2.005376],accel_mss,speed_ms,0,blend_radius_m)
  movel([0.431281, -0.497135, -2.827313, -1.387941, 1.570796, 2.002077],accel_mss,speed_ms,0,blend_radius_m)
  movel([0.427645, -0.504914, -2.826979, -1.380496, 1.570796, 1.998441],accel_mss,speed_ms,0,blend_radius_m)
  movel([0.423704, -0.512789, -2.826619, -1.372981, 1.570796, 1.994500],accel_mss,speed_ms,0,blend_radius_m)
  movel([0.419475, -0.520714, -2.826235, -1.365440, 1.570796, 1.990272],accel_mss,speed_ms,0,blend_radius_m)
  movel([0.414991, -0.528655, -2.825827, -1.357906, 1.570796, 1.985787],accel_mss,speed_ms,0,blend_radius_m)
  movel([0.410254, -0.536589, -2.825397, -1.350403, 1.570796, 1.981050],accel_mss,speed_ms,0,blend_radius_m)
  movel([0.405294, -0.544482, -2.824947, -1.342960, 1.570796, 1.976090],accel_mss,speed_ms,0,blend_radius_m)
  movel([0.401988, -0.549431, -2.824653, -1.338305, 1.570796, 1.972784],accel_mss,speed_ms,0,blend_radius_m)
  movel([0.398403, -0.554269, -2.824357, -1.333763, 1.570796, 1.969199],accel_mss,speed_ms,0,blend_radius_m)
  movel([0.394613, -0.558623, -2.824083, -1.329683, 1.570796, 1.965409],accel_mss,speed_ms,0,blend_radius_m)
  movel([0.392667, -0.560491, -2.823963, -1.327934, 1.570796, 1.963463],accel_mss,speed_ms,0,blend_radius_m)
  movel([0.390691, -0.562108, -2.823859, -1.326422, 1.570796, 1.961488],accel_mss,speed_ms,0,blend_radius_m)
  speed_ms = 0.005
  movel([0.390691, -0.557222, -2.816971, -1.338196, 1.570796, 1.961488],accel_mss,speed_ms,0,blend_radius_m)
  speed_ms = 0.040
  movel([0.379771, -0.570764, -2.816059, -1.325566, 1.570796, 1.950568],accel_mss,speed_ms,0,blend_radius_m)
  speed_ms = 0.005
  movel([0.379771, -0.575892, -2.822928, -1.313569, 1.570796, 1.950568],accel_mss,speed_ms,0,blend_radius_m)
  speed_ms = 0.025
  movel([0.379949, -0.576942, -2.822854, -1.312593, 1.570796, 1.950745],accel_mss,speed_ms,0,blend_radius_m)
  movel([0.379468, -0.578533, -2.822741, -1.311114, 1.570796, 1.950264],accel_mss,speed_ms,0,blend_radius_m)
  movel([0.378499, -0.580394, -2.822608, -1.309386, 1.570796, 1.949295],accel_mss,speed_ms,0,blend_radius_m)
  movel([0.377199, -0.582254, -2.822474, -1.307661, 1.570796, 1.947995],accel_mss,speed_ms,0,blend_radius_m)
  movel([0.375432, -0.584139, -2.822337, -1.305913, 1.570796, 1.946228],accel_mss,speed_ms,0,blend_radius_m)
  movel([0.373657, -0.585636, -2.822227, -1.304526, 1.570796, 1.944453],accel_mss,speed_ms,0,blend_radius_m)
  movel([0.371926, -0.587038, -2.822123, -1.303228, 1.570796, 1.942722],accel_mss,speed_ms,0,blend_radius_m)
  movel([0.370313, -0.588638, -2.822003, -1.301747, 1.570796, 1.941109],accel_mss,speed_ms,0,blend_radius_m)
  movel([0.368536, -0.591344, -2.821799, -1.299246, 1.570796, 1.939332],accel_mss,speed_ms,0,blend_radius_m)
  movel([0.367706, -0.592751, -2.821692, -1.297946, 1.570796, 1.938503],accel_mss,speed_ms,0,blend_radius_m)
  movel([0.366616, -0.594243, -2.821577, -1.296568, 1.570796, 1.937412],accel_mss,speed_ms,0,blend_radius_m)
  movel([0.363281, -0.597945, -2.821289, -1.293155, 1.570796, 1.934078],accel_mss,speed_ms,0,blend_radius_m)
  movel([0.359964, -0.601129, -2.821037, -1.290223, 1.570796, 1.930761],accel_mss,speed_ms,0,blend_radius_m)
  movel([0.356635, -0.603873, -2.820817, -1.287699, 1.570796, 1.927431],accel_mss,speed_ms,0,blend_radius_m)
  movel([0.353259, -0.606285, -2.820621, -1.285483, 1.570796, 1.924055],accel_mss,speed_ms,0,blend_radius_m)
  movel([0.355034, -0.604852, -2.820738, -1.286799, 1.570796, 1.925830],accel_mss,speed_ms,0,blend_radius_m)
  movel([0.356757, -0.603698, -2.820831, -1.287860, 1.570796, 1.927553],accel_mss,speed_ms,0,blend_radius_m)
  movel([0.358252, -0.603188, -2.820872, -1.288328, 1.570796, 1.929048],accel_mss,speed_ms,0,blend_radius_m)
  movel([0.359104, -0.603683, -2.820832, -1.287874, 1.570796, 1.929901],accel_mss,speed_ms,0,blend_radius_m)
  movel([0.358949, -0.605203, -2.820709, -1.286477, 1.570796, 1.929745],accel_mss,speed_ms,0,blend_radius_m)
  movel([0.358015, -0.607198, -2.820546, -1.284645, 1.570796, 1.928811],accel_mss,speed_ms,0,blend_radius_m)
  movel([0.356611, -0.609221, -2.820379, -1.282789, 1.570796, 1.927407],accel_mss,speed_ms,0,blend_radius_m)
  movel([0.352353, -0.614033, -2.819976, -1.278380, 1.570796, 1.923149],accel_mss,speed_ms,0,blend_radius_m)
  movel([0.349628, -0.616694, -2.819749, -1.275947, 1.570796, 1.920424],accel_mss,speed_ms,0,blend_radius_m)
  movel([0.346894, -0.619076, -2.819543, -1.273770, 1.570796, 1.917690],accel_mss,speed_ms,0,blend_radius_m)
  movel([0.344176, -0.621151, -2.819362, -1.271876, 1.570796, 1.914972],accel_mss,speed_ms,0,blend_radius_m)
  movel([0.347204, -0.619232, -2.819530, -1.273627, 1.570796, 1.918001],accel_mss,speed_ms,0,blend_radius_m)
  movel([0.350417, -0.616841, -2.819736, -1.275812, 1.570796, 1.921214],accel_mss,speed_ms,0,blend_radius_m)
  movel([0.353558, -0.614567, -2.819930, -1.277892, 1.570796, 1.924354],accel_mss,speed_ms,0,blend_radius_m)
  movel([0.356373, -0.612974, -2.820065, -1.279350, 1.570796, 1.927169],accel_mss,speed_ms,0,blend_radius_m)
  movel([0.357104, -0.612900, -2.820072, -1.279417, 1.570796, 1.927900],accel_mss,speed_ms,0,blend_radius_m)
  movel([0.357042, -0.613516, -2.820020, -1.278854, 1.570796, 1.927838],accel_mss,speed_ms,0,blend_radius_m)
  movel([0.355138, -0.616812, -2.819739, -1.275838, 1.570796, 1.925934],accel_mss,speed_ms,0,blend_radius_m)
  movel([0.353460, -0.619205, -2.819532, -1.273652, 1.570796, 1.924257],accel_mss,speed_ms,0,blend_radius_m)
  movel([0.351629, -0.621502, -2.819332, -1.271556, 1.570796, 1.922426],accel_mss,speed_ms,0,blend_radius_m)
  movel([0.349693, -0.623640, -2.819143, -1.269606, 1.570796, 1.920490],accel_mss,speed_ms,0,blend_radius_m)
  movel([0.350644, -0.622808, -2.819217, -1.270364, 1.570796, 1.921441],accel_mss,speed_ms,0,blend_radius_m)
  movel([0.351670, -0.622177, -2.819272, -1.270940, 1.570796, 1.922466],accel_mss,speed_ms,0,blend_radius_m)
  movel([0.353820, -0.621465, -2.819335, -1.271590, 1.570796, 1.924616],accel_mss,speed_ms,0,blend_radius_m)
  movel([0.355869, -0.621432, -2.819338, -1.271619, 1.570796, 1.926665],accel_mss,speed_ms,0,blend_radius_m)
  movel([0.357562, -0.621994, -2.819288, -1.271107, 1.570796, 1.928358],accel_mss,speed_ms,0,blend_radius_m)
  movel([0.358648, -0.623060, -2.819194, -1.270135, 1.570796, 1.929444],accel_mss,speed_ms,0,blend_radius_m)
  movel([0.358876, -0.624532, -2.819064, -1.268793, 1.570796, 1.929673],accel_mss,speed_ms,0,blend_radius_m)
  movel([0.358591, -0.625391, -2.818987, -1.268011, 1.570796, 1.929388],accel_mss,speed_ms,0,blend_radius_m)
  movel([0.357999, -0.626312, -2.818905, -1.267172, 1.570796, 1.928795],accel_mss,speed_ms,0,blend_radius_m)
  movel([0.357072, -0.627295, -2.818817, -1.266278, 1.570796, 1.927869],accel_mss,speed_ms,0,blend_radius_m)
  movel([0.355773, -0.628318, -2.818724, -1.265346, 1.570796, 1.926569],accel_mss,speed_ms,0,blend_radius_m)
  movel([0.354385, -0.629056, -2.818657, -1.264676, 1.570796, 1.925181],accel_mss,speed_ms,0,blend_radius_m)
  movel([0.349446, -0.629892, -2.818581, -1.263915, 1.570796, 1.920242],accel_mss,speed_ms,0,blend_radius_m)
  movel([0.347504, -0.630348, -2.818540, -1.263501, 1.570796, 1.918301],accel_mss,speed_ms,0,blend_radius_m)
  movel([0.345366, -0.631265, -2.818456, -1.262668, 1.570796, 1.916163],accel_mss,speed_ms,0,blend_radius_m)
  movel([0.341503, -0.633866, -2.818216, -1.260306, 1.570796, 1.912300],accel_mss,speed_ms,0,blend_radius_m)
  movel([0.337576, -0.636763, -2.817946, -1.257680, 1.570796, 1.908372],accel_mss,speed_ms,0,blend_radius_m)
  movel([0.335660, -0.637879, -2.817841, -1.256669, 1.570796, 1.906456],accel_mss,speed_ms,0,blend_radius_m)
  movel([0.333925, -0.638513, -2.817781, -1.256095, 1.570796, 1.904721],accel_mss,speed_ms,0,blend_radius_m)
  movel([0.332602, -0.638475, -2.817785, -1.256129, 1.570796, 1.903398],accel_mss,speed_ms,0,blend_radius_m)
  movel([0.331912, -0.637587, -2.817869, -1.256933, 1.570796, 1.902709],accel_mss,speed_ms,0,blend_radius_m)
  movel([0.333990, -0.634858, -2.818124, -1.259407, 1.570796, 1.904787],accel_mss,speed_ms,0,blend_radius_m)
  movel([0.336211, -0.632253, -2.818365, -1.261771, 1.570796, 1.907007],accel_mss,speed_ms,0,blend_radius_m)
  speed_ms = 0.005
  movel([0.336211, -0.626188, -2.811588, -1.274613, 1.570796, 1.907007],accel_mss,speed_ms,0,blend_radius_m)
  speed_ms = 0.040
  movel([0.351549, -0.635617, -2.810706, -1.266067, 1.570796, 1.922345],accel_mss,speed_ms,0,blend_radius_m)
  speed_ms = 0.005
  movel([0.351549, -0.641832, -2.817465, -1.253091, 1.570796, 1.922345],accel_mss,speed_ms,0,blend_radius_m)
  speed_ms = 0.025
  movel([0.353017, -0.639886, -2.817651, -1.254852, 1.570796, 1.923813],accel_mss,speed_ms,0,blend_radius_m)
  movel([0.354736, -0.638395, -2.817792, -1.256201, 1.570796, 1.925532],accel_mss,speed_ms,0,blend_radius_m)
  movel([0.356426, -0.637488, -2.817878, -1.257023, 1.570796, 1.927223],accel_mss,speed_ms,0,blend_radius_m)
  movel([0.357799, -0.637301, -2.817896, -1.257193, 1.570796, 1.928595],accel_mss,speed_ms,0,blend_radius_m)
  movel([0.358713, -0.637784, -2.817850, -1.256755, 1.570796, 1.929509],accel_mss,speed_ms,0,blend_radius_m)
  movel([0.359289, -0.638695, -2.817764, -1.255930, 1.570796, 1.930085],accel_mss,speed_ms,0,blend_radius_m)
  movel([0.359851, -0.641190, -2.817527, -1.253672, 1.570796, 1.930648],accel_mss,speed_ms,0,blend_radius_m)
  movel([0.361230, -0.638814, -2.817753, -1.255822, 1.570796, 1.932027],accel_mss,speed_ms,0,blend_radius_m)
  movel([0.362162, -0.636531, -2.817968, -1.257890, 1.570796, 1.932958],accel_mss,speed_ms,0,blend_radius_m)
  movel([0.362570, -0.634541, -2.818154, -1.259694, 1.570796, 1.933367],accel_mss,speed_ms,0,blend_radius_m)
  movel([0.362409, -0.633006, -2.818296, -1.261087, 1.570796, 1.933205],accel_mss,speed_ms,0,blend_radius_m)
  movel([0.363247, -0.633431, -2.818257, -1.260702, 1.570796, 1.934044],accel_mss,speed_ms,0,blend_radius_m)
  movel([0.363803, -0.634191, -2.818186, -1.260012, 1.570796, 1.934599],accel_mss,speed_ms,0,blend_radius_m)
  movel([0.364218, -0.636485, -2.817972, -1.257932, 1.570796, 1.935014],accel_mss,speed_ms,0,blend_radius_m)
  movel([0.363986, -0.639449, -2.817693, -1.255248, 1.570796, 1.934783],accel_mss,speed_ms,0,blend_radius_m)
  movel([0.363403, -0.642676, -2.817384, -1.252328, 1.570796, 1.934200],accel_mss,speed_ms,0,blend_radius_m)
  movel([0.362304, -0.646445, -2.817018, -1.248926, 1.570796, 1.933101],accel_mss,speed_ms,0,blend_radius_m)
  movel([0.360800, -0.650209, -2.816648, -1.245533, 1.570796, 1.931596],accel_mss,speed_ms,0,blend_radius_m)
  movel([0.359255, -0.653922, -2.816276, -1.242191, 1.570796, 1.930051],accel_mss,speed_ms,0,blend_radius_m)
  movel([0.358028, -0.657552, -2.815907, -1.238930, 1.570796, 1.928824],accel_mss,speed_ms,0,blend_radius_m)
  movel([0.357067, -0.655954, -2.816070, -1.240365, 1.570796, 1.927863],accel_mss,speed_ms,0,blend_radius_m)
  movel([0.355532, -0.655088, -2.816158, -1.241143, 1.570796, 1.926329],accel_mss,speed_ms,0,blend_radius_m)
  movel([0.353464, -0.655028, -2.816164, -1.241197, 1.570796, 1.924261],accel_mss,speed_ms,0,blend_radius_m)
  movel([0.350894, -0.655853, -2.816080, -1.240456, 1.570796, 1.921690],accel_mss,speed_ms,0,blend_radius_m)
  speed_ms = 0.005
  movel([0.350894, -0.649422, -2.809348, -1.253620, 1.570796, 1.921690],accel_mss,speed_ms,0,blend_radius_m)
  speed_ms = 0.040
  movel([0.352138, -0.658896, -2.808370, -1.245123, 1.570796, 1.922935],accel_mss,speed_ms,0,blend_radius_m)
  speed_ms = 0.005
  movel([0.352138, -0.665472, -2.815083, -1.231834, 1.570796, 1.922935],accel_mss,speed_ms,0,blend_radius_m)
  speed_ms = 0.025
  movel([0.351964, -0.669567, -2.814647, -1.228175, 1.570796, 1.922760],accel_mss,speed_ms,0,blend_radius_m)
  movel([0.352428, -0.673096, -2.814265, -1.225028, 1.570796, 1.923224],accel_mss,speed_ms,0,blend_radius_m)
  movel([0.353764, -0.675630, -2.813988, -1.222771, 1.570796, 1.924560],accel_mss,speed_ms,0,blend_radius_m)
  movel([0.354836, -0.676390, -2.813904, -1.222095, 1.570796, 1.925632],accel_mss,speed_ms,0,blend_radius_m)
  movel([0.356219, -0.676743, -2.813865, -1.221781, 1.570796, 1.927016],accel_mss,speed_ms,0,blend_radius_m)
  movel([0.358558, -0.676499, -2.813892, -1.221998, 1.570796, 1.929355],accel_mss,speed_ms,0,blend_radius_m)
  movel([0.361206, -0.675537, -2.813998, -1.222853, 1.570796, 1.932002],accel_mss,speed_ms,0,blend_radius_m)
  movel([0.364101, -0.674023, -2.814164, -1.224202, 1.570796, 1.934897],accel_mss,speed_ms,0,blend_radius_m)
  movel([0.367174, -0.672121, -2.814371, -1.225897, 1.570796, 1.937971],accel_mss,speed_ms,0,blend_radius_m)
  movel([0.373586, -0.667806, -2.814835, -1.229748, 1.570796, 1.944382],accel_mss,speed_ms,0,blend_radius_m)
  movel([0.379870, -0.663942, -2.815244, -1.233203, 1.570796, 1.950666],accel_mss,speed_ms,0,blend_radius_m)
  movel([0.383258, -0.662419, -2.815404, -1.234567, 1.570796, 1.954054],accel_mss,speed_ms,0,blend_radius_m)
  movel([0.386363, -0.661562, -2.815493, -1.235334, 1.570796, 1.957160],accel_mss,speed_ms,0,blend_radius_m)
  movel([0.389136, -0.661357, -2.815515, -1.235518, 1.570796, 1.959932],accel_mss,speed_ms,0,blend_radius_m)
  movel([0.391521, -0.661797, -2.815469, -1.235124, 1.570796, 1.962317],accel_mss,speed_ms,0,blend_radius_m)
  movel([0.393479, -0.662853, -2.815359, -1.234178, 1.570796, 1.964275],accel_mss,speed_ms,0,blend_radius_m)
  movel([0.394959, -0.664514, -2.815184, -1.232690, 1.570796, 1.965755],accel_mss,speed_ms,0,blend_radius_m)
  movel([0.395914, -0.666759, -2.814947, -1.230683, 1.570796, 1.966710],accel_mss,speed_ms,0,blend_radius_m)
  movel([0.396312, -0.669555, -2.814648, -1.228186, 1.570796, 1.967108],accel_mss,speed_ms,0,blend_radius_m)
  speed_ms = 0.005
  movel([0.396312, -0.662918, -2.807944, -1.241528, 1.570796, 1.967108],accel_mss,speed_ms,0,blend_radius_m)
  speed_ms = 0.040
  movel([0.345905, -0.631067, -2.811136, -1.270186, 1.570796, 1.916701],accel_mss,speed_ms,0,blend_radius_m)
  speed_ms = 0.005
  movel([0.345905, -0.637211, -2.817904, -1.257274, 1.570796, 1.916701],accel_mss,speed_ms,0,blend_radius_m)
  speed_ms = 0.025
  movel([0.347293, -0.637524, -2.817875, -1.256991, 1.570796, 1.918089],accel_mss,speed_ms,0,blend_radius_m)
  movel([0.348210, -0.638439, -2.817788, -1.256162, 1.570796, 1.919007],accel_mss,speed_ms,0,blend_radius_m)
  movel([0.348304, -0.639300, -2.817707, -1.255382, 1.570796, 1.919100],accel_mss,speed_ms,0,blend_radius_m)
  movel([0.348070, -0.640424, -2.817600, -1.254365, 1.570796, 1.918866],accel_mss,speed_ms,0,blend_radius_m)
  movel([0.347517, -0.641684, -2.817479, -1.253226, 1.570796, 1.918313],accel_mss,speed_ms,0,blend_radius_m)
  movel([0.346644, -0.642957, -2.817357, -1.252075, 1.570796, 1.917440],accel_mss,speed_ms,0,blend_radius_m)
  movel([0.344727, -0.645066, -2.817153, -1.250170, 1.570796, 1.915523],accel_mss,speed_ms,0,blend_radius_m)
  movel([0.343988, -0.646269, -2.817036, -1.249084, 1.570796, 1.914784],accel_mss,speed_ms,0,blend_radius_m)
  movel([0.343592, -0.647403, -2.816925, -1.248061, 1.570796, 1.914388],accel_mss,speed_ms,0,blend_radius_m)
  movel([0.343551, -0.649274, -2.816740, -1.246375, 1.570796, 1.914347],accel_mss,speed_ms,0,blend_radius_m)
  movel([0.344108, -0.650902, -2.816579, -1.244909, 1.570796, 1.914905],accel_mss,speed_ms,0,blend_radius_m)
  movel([0.345022, -0.652131, -2.816456, -1.243802, 1.570796, 1.915818],accel_mss,speed_ms,0,blend_radius_m)
  movel([0.346266, -0.652956, -2.816373, -1.243060, 1.570796, 1.917062],accel_mss,speed_ms,0,blend_radius_m)
  movel([0.347814, -0.653348, -2.816334, -1.242707, 1.570796, 1.918611],accel_mss,speed_ms,0,blend_radius_m)
  movel([0.346143, -0.656038, -2.816062, -1.240290, 1.570796, 1.916940],accel_mss,speed_ms,0,blend_radius_m)
  movel([0.344813, -0.658653, -2.815794, -1.237942, 1.570796, 1.915609],accel_mss,speed_ms,0,blend_radius_m)
  movel([0.343783, -0.661190, -2.815532, -1.235667, 1.570796, 1.914580],accel_mss,speed_ms,0,blend_radius_m)
  movel([0.343015, -0.663638, -2.815276, -1.233475, 1.570796, 1.913812],accel_mss,speed_ms,0,blend_radius_m)
  movel([0.342123, -0.668235, -2.814790, -1.229365, 1.570796, 1.912920],accel_mss,speed_ms,0,blend_radius_m)
  movel([0.341863, -0.672371, -2.814344, -1.225674, 1.570796, 1.912659],accel_mss,speed_ms,0,blend_radius_m)
  movel([0.341691, -0.676301, -2.813914, -1.222174, 1.570796, 1.912487],accel_mss,speed_ms,0,blend_radius_m)
  movel([0.341301, -0.678458, -2.813675, -1.220256, 1.570796, 1.912097],accel_mss,speed_ms,0,blend_radius_m)
  movel([0.340520, -0.680831, -2.813410, -1.218147, 1.570796, 1.911316],accel_mss,speed_ms,0,blend_radius_m)
  movel([0.339172, -0.683442, -2.813116, -1.215831, 1.570796, 1.909969],accel_mss,speed_ms,0,blend_radius_m)
  movel([0.337350, -0.685999, -2.812825, -1.213565, 1.570796, 1.908147],accel_mss,speed_ms,0,blend_radius_m)
  movel([0.335304, -0.688105, -2.812583, -1.211701, 1.570796, 1.906101],accel_mss,speed_ms,0,blend_radius_m)
  movel([0.333296, -0.689350, -2.812439, -1.210601, 1.570796, 1.904092],accel_mss,speed_ms,0,blend_radius_m)
  movel([0.333851, -0.690663, -2.812286, -1.209439, 1.570796, 1.904647],accel_mss,speed_ms,0,blend_radius_m)
  movel([0.334133, -0.694075, -2.811887, -1.206427, 1.570796, 1.904930],accel_mss,speed_ms,0,blend_radius_m)
  movel([0.333871, -0.696105, -2.811646, -1.204638, 1.570796, 1.904667],accel_mss,speed_ms,0,blend_radius_m)
  movel([0.332594, -0.700621, -2.811105, -1.200663, 1.570796, 1.903390],accel_mss,speed_ms,0,blend_radius_m)
  movel([0.331591, -0.703034, -2.810812, -1.198543, 1.570796, 1.902387],accel_mss,speed_ms,0,blend_radius_m)
  movel([0.330351, -0.705510, -2.810509, -1.196370, 1.570796, 1.901147],accel_mss,speed_ms,0,blend_radius_m)
  speed_ms = 0.005
  movel([0.330351, -0.698361, -2.803884, -1.210144, 1.570796, 1.901147],accel_mss,speed_ms,0,blend_radius_m)
  speed_ms = 0.040
  movel([0.320831, -0.702434, -2.803382, -1.206573, 1.570796, 1.891628],accel_mss,speed_ms,0,blend_radius_m)
  speed_ms = 0.005
  movel([0.320831, -0.709639, -2.809998, -1.192752, 1.570796, 1.891628],accel_mss,speed_ms,0,blend_radius_m)
  speed_ms = 0.025
  movel([0.323413, -0.726531, -2.807825, -1.178033, 1.570796, 1.894209],accel_mss,speed_ms,0,blend_radius_m)
  movel([0.323461, -0.728810, -2.807522, -1.176057, 1.570796, 1.894258],accel_mss,speed_ms,0,blend_radius_m)
  movel([0.323113, -0.730145, -2.807343, -1.174901, 1.570796, 1.893909],accel_mss,speed_ms,0,blend_radius_m)
  movel([0.322352, -0.731599, -2.807148, -1.173642, 1.570796, 1.893148],accel_mss,speed_ms,0,blend_radius_m)
  movel([0.320056, -0.734673, -2.806731, -1.170985, 1.570796, 1.890852],accel_mss,speed_ms,0,blend_radius_m)
  movel([0.319501, -0.736192, -2.806524, -1.169673, 1.570796, 1.890297],accel_mss,speed_ms,0,blend_radius_m)
  movel([0.319482, -0.737433, -2.806353, -1.168603, 1.570796, 1.890279],accel_mss,speed_ms,0,blend_radius_m)
  movel([0.320112, -0.738923, -2.806148, -1.167318, 1.570796, 1.890908],accel_mss,speed_ms,0,blend_radius_m)
  movel([0.321291, -0.739887, -2.806014, -1.166487, 1.570796, 1.892088],accel_mss,speed_ms,0,blend_radius_m)
  movel([0.323990, -0.741286, -2.805820, -1.165283, 1.570796, 1.894786],accel_mss,speed_ms,0,blend_radius_m)
  movel([0.325329, -0.742762, -2.805614, -1.164013, 1.570796, 1.896125],accel_mss,speed_ms,0,blend_radius_m)
  movel([0.326698, -0.745424, -2.805239, -1.161726, 1.570796, 1.897494],accel_mss,speed_ms,0,blend_radius_m)
  movel([0.326968, -0.746939, -2.805025, -1.160426, 1.570796, 1.897764],accel_mss,speed_ms,0,blend_radius_m)
  movel([0.326754, -0.748426, -2.804813, -1.159150, 1.570796, 1.897550],accel_mss,speed_ms,0,blend_radius_m)
  movel([0.326410, -0.749125, -2.804713, -1.158551, 1.570796, 1.897207],accel_mss,speed_ms,0,blend_radius_m)
  movel([0.325881, -0.749775, -2.804620, -1.157994, 1.570796, 1.896678],accel_mss,speed_ms,0,blend_radius_m)
  movel([0.324184, -0.750893, -2.804460, -1.157036, 1.570796, 1.894981],accel_mss,speed_ms,0,blend_radius_m)
  movel([0.324146, -0.752370, -2.804247, -1.155773, 1.570796, 1.894943],accel_mss,speed_ms,0,blend_radius_m)
  movel([0.324547, -0.753706, -2.804053, -1.154630, 1.570796, 1.895344],accel_mss,speed_ms,0,blend_radius_m)
  movel([0.326252, -0.755952, -2.803726, -1.152711, 1.570796, 1.897049],accel_mss,speed_ms,0,blend_radius_m)
  movel([0.330428, -0.758817, -2.803305, -1.150267, 1.570796, 1.901225],accel_mss,speed_ms,0,blend_radius_m)
  movel([0.332973, -0.759602, -2.803189, -1.149599, 1.570796, 1.903769],accel_mss,speed_ms,0,blend_radius_m)
  movel([0.335888, -0.760049, -2.803122, -1.149218, 1.570796, 1.906684],accel_mss,speed_ms,0,blend_radius_m)
  movel([0.338411, -0.760970, -2.802985, -1.148433, 1.570796, 1.909207],accel_mss,speed_ms,0,blend_radius_m)
  movel([0.339288, -0.761856, -2.802854, -1.147680, 1.570796, 1.910085],accel_mss,speed_ms,0,blend_radius_m)
  movel([0.339784, -0.763158, -2.802659, -1.146572, 1.570796, 1.910580],accel_mss,speed_ms,0,blend_radius_m)
  movel([0.339779, -0.764062, -2.802523, -1.145804, 1.570796, 1.910575],accel_mss,speed_ms,0,blend_radius_m)
  movel([0.339496, -0.765137, -2.802362, -1.144891, 1.570796, 1.910293],accel_mss,speed_ms,0,blend_radius_m)
  movel([0.338944, -0.766189, -2.802203, -1.143997, 1.570796, 1.909740],accel_mss,speed_ms,0,blend_radius_m)
  movel([0.338115, -0.767024, -2.802076, -1.143289, 1.570796, 1.908911],accel_mss,speed_ms,0,blend_radius_m)
  movel([0.336844, -0.767356, -2.802026, -1.143007, 1.570796, 1.907640],accel_mss,speed_ms,0,blend_radius_m)
  movel([0.331845, -0.766678, -2.802129, -1.143582, 1.570796, 1.902641],accel_mss,speed_ms,0,blend_radius_m)
  movel([0.327463, -0.765048, -2.802375, -1.144966, 1.570796, 1.898259],accel_mss,speed_ms,0,blend_radius_m)
  movel([0.326911, -0.766235, -2.802196, -1.143958, 1.570796, 1.897708],accel_mss,speed_ms,0,blend_radius_m)
  movel([0.326609, -0.767331, -2.802030, -1.143029, 1.570796, 1.897405],accel_mss,speed_ms,0,blend_radius_m)
  movel([0.326653, -0.769262, -2.801736, -1.141392, 1.570796, 1.897450],accel_mss,speed_ms,0,blend_radius_m)
  movel([0.327394, -0.770865, -2.801490, -1.140034, 1.570796, 1.898190],accel_mss,speed_ms,0,blend_radius_m)
  movel([0.328616, -0.772195, -2.801285, -1.138909, 1.570796, 1.899412],accel_mss,speed_ms,0,blend_radius_m)
  movel([0.331744, -0.774116, -2.800988, -1.137285, 1.570796, 1.902540],accel_mss,speed_ms,0,blend_radius_m)
  movel([0.334451, -0.775270, -2.800809, -1.136311, 1.570796, 1.905247],accel_mss,speed_ms,0,blend_radius_m)
  movel([0.335324, -0.775870, -2.800715, -1.135804, 1.570796, 1.906121],accel_mss,speed_ms,0,blend_radius_m)
  movel([0.335511, -0.776407, -2.800631, -1.135350, 1.570796, 1.906307],accel_mss,speed_ms,0,blend_radius_m)
  movel([0.335387, -0.777181, -2.800510, -1.134698, 1.570796, 1.906183],accel_mss,speed_ms,0,blend_radius_m)
  movel([0.334923, -0.778144, -2.800359, -1.133886, 1.570796, 1.905720],accel_mss,speed_ms,0,blend_radius_m)
  movel([0.334354, -0.778841, -2.800250, -1.133299, 1.570796, 1.905150],accel_mss,speed_ms,0,blend_radius_m)
  movel([0.333034, -0.779710, -2.800112, -1.132566, 1.570796, 1.903831],accel_mss,speed_ms,0,blend_radius_m)
  movel([0.331203, -0.780728, -2.799951, -1.131710, 1.570796, 1.901999],accel_mss,speed_ms,0,blend_radius_m)
  movel([0.330790, -0.781259, -2.799867, -1.131263, 1.570796, 1.901586],accel_mss,speed_ms,0,blend_radius_m)
  movel([0.330501, -0.782054, -2.799741, -1.130594, 1.570796, 1.901297],accel_mss,speed_ms,0,blend_radius_m)
  movel([0.330491, -0.782781, -2.799625, -1.129983, 1.570796, 1.901287],accel_mss,speed_ms,0,blend_radius_m)
  movel([0.331058, -0.784017, -2.799427, -1.128944, 1.570796, 1.901854],accel_mss,speed_ms,0,blend_radius_m)
  movel([0.332754, -0.785671, -2.799162, -1.127556, 1.570796, 1.903551],accel_mss,speed_ms,0,blend_radius_m)
  movel([0.340812, -0.791597, -2.798199, -1.122593, 1.570796, 1.911608],accel_mss,speed_ms,0,blend_radius_m)
  movel([0.341451, -0.792403, -2.798067, -1.121919, 1.570796, 1.912247],accel_mss,speed_ms,0,blend_radius_m)
  movel([0.341793, -0.793511, -2.797884, -1.120993, 1.570796, 1.912589],accel_mss,speed_ms,0,blend_radius_m)
  movel([0.341637, -0.794880, -2.797658, -1.119850, 1.570796, 1.912433],accel_mss,speed_ms,0,blend_radius_m)
  movel([0.340781, -0.796459, -2.797396, -1.118534, 1.570796, 1.911578],accel_mss,speed_ms,0,blend_radius_m)
